(* IEC 61131-3 sources: BODAS-RC27-18_40/st/bodas_rc18_12_27_18_40/plc_logic/application/dsm_easyconfig/structure (part 2) *)

(* ---- dfc_rbr_ina57or-DFC_rbr_inA57OR.st ---- *)
(* --- Interface --- *)
{attribute 'external_name' := 'cmp_rts_DFC_rbr_inA57OR'}
TYPE DFC_rbr_inA57OR :
STRUCT
	DTC: UDINT := 16#134C00;
	DFCid: UINT := 81;
	debounceMethod: USINT := TIME_UP_DOWN;
END_STRUCT
END_TYPE

(* ---- dfc_rbr_ina57scb-DFC_rbr_inA57SCB.st ---- *)
(* --- Interface --- *)
{attribute 'external_name' := 'cmp_rts_DFC_rbr_inA57SCB'}
TYPE DFC_rbr_inA57SCB :
STRUCT
	DTC: UDINT := 16#134D00;
	DFCid: UINT := 82;
	debounceMethod: USINT := TIME_UP_DOWN;
END_STRUCT
END_TYPE

(* ---- dfc_rbr_ina57scg-DFC_rbr_inA57SCG.st ---- *)
(* --- Interface --- *)
{attribute 'external_name' := 'cmp_rts_DFC_rbr_inA57SCG'}
TYPE DFC_rbr_inA57SCG :
STRUCT
	DTC: UDINT := 16#134E00;
	DFCid: UINT := 83;
	debounceMethod: USINT := TIME_UP_DOWN;
END_STRUCT
END_TYPE

(* ---- dfc_rbr_ina59ol-DFC_rbr_inA59OL.st ---- *)
(* --- Interface --- *)
{attribute 'external_name' := 'cmp_rts_DFC_rbr_inA59OL'}
TYPE DFC_rbr_inA59OL :
STRUCT
	DTC: UDINT := 16#134F00;
	DFCid: UINT := 84;
	debounceMethod: USINT := TIME_UP_DOWN;
END_STRUCT
END_TYPE

(* ---- dfc_rbr_ina59scb-DFC_rbr_inA59SCB.st ---- *)
(* --- Interface --- *)
{attribute 'external_name' := 'cmp_rts_DFC_rbr_inA59SCB'}
TYPE DFC_rbr_inA59SCB :
STRUCT
	DTC: UDINT := 16#135000;
	DFCid: UINT := 85;
	debounceMethod: USINT := TIME_UP_DOWN;
END_STRUCT
END_TYPE

(* ---- dfc_rbr_ina59scg-DFC_rbr_inA59SCG.st ---- *)
(* --- Interface --- *)
{attribute 'external_name' := 'cmp_rts_DFC_rbr_inA59SCG'}
TYPE DFC_rbr_inA59SCG :
STRUCT
	DTC: UDINT := 16#135100;
	DFCid: UINT := 86;
	debounceMethod: USINT := TIME_UP_DOWN;
END_STRUCT
END_TYPE

(* ---- dfc_rbr_inai-DFC_rbr_inAi.st ---- *)
(* --- Interface --- *)
{attribute 'external_name' := 'cmp_rts_DFC_rbr_inAi'}
TYPE DFC_rbr_inAi :
STRUCT
	DTC: UDINT := 16#038000;
	DFCid: UINT := 578;
	debounceMethod: USINT := NO_DEBOUNCE;
END_STRUCT
END_TYPE

(* ---- dfc_rbr_inaic-DFC_rbr_inAic.st ---- *)
(* --- Interface --- *)
{attribute 'external_name' := 'cmp_rts_DFC_rbr_inAic'}
TYPE DFC_rbr_inAic :
STRUCT
	DTC: UDINT := 16#038100;
	DFCid: UINT := 579;
	debounceMethod: USINT := NO_DEBOUNCE;
END_STRUCT
END_TYPE

(* ---- dfc_rbr_inaiccfg-DFC_rbr_inAicCfg.st ---- *)
(* --- Interface --- *)
{attribute 'external_name' := 'cmp_rts_DFC_rbr_inAicCfg'}
TYPE DFC_rbr_inAicCfg :
STRUCT
	DTC: UDINT := 16#038200;
	DFCid: UINT := 580;
	debounceMethod: USINT := NO_DEBOUNCE;
END_STRUCT
END_TYPE

(* ---- dfc_rbr_inaicgetstatus-DFC_rbr_inAicGetStatus.st ---- *)
(* --- Interface --- *)
{attribute 'external_name' := 'cmp_rts_DFC_rbr_inAicGetStatus'}
TYPE DFC_rbr_inAicGetStatus :
STRUCT
	DTC: UDINT := 16#038D00;
	DFCid: UINT := 581;
	debounceMethod: USINT := NO_DEBOUNCE;
END_STRUCT
END_TYPE

(* ---- dfc_rbr_inaid-DFC_rbr_inAid.st ---- *)
(* --- Interface --- *)
{attribute 'external_name' := 'cmp_rts_DFC_rbr_inAid'}
TYPE DFC_rbr_inAid :
STRUCT
	DTC: UDINT := 16#038300;
	DFCid: UINT := 582;
	debounceMethod: USINT := NO_DEBOUNCE;
END_STRUCT
END_TYPE

(* ---- dfc_rbr_inaidcfg-DFC_rbr_inAidCfg.st ---- *)
(* --- Interface --- *)
{attribute 'external_name' := 'cmp_rts_DFC_rbr_inAidCfg'}
TYPE DFC_rbr_inAidCfg :
STRUCT
	DTC: UDINT := 16#038400;
	DFCid: UINT := 583;
	debounceMethod: USINT := NO_DEBOUNCE;
END_STRUCT
END_TYPE

(* ---- dfc_rbr_inaiv-DFC_rbr_inAiv.st ---- *)
(* --- Interface --- *)
{attribute 'external_name' := 'cmp_rts_DFC_rbr_inAiv'}
TYPE DFC_rbr_inAiv :
STRUCT
	DTC: UDINT := 16#038500;
	DFCid: UINT := 584;
	debounceMethod: USINT := NO_DEBOUNCE;
END_STRUCT
END_TYPE

(* ---- dfc_rbr_inaivcfg-DFC_rbr_inAivCfg.st ---- *)
(* --- Interface --- *)
{attribute 'external_name' := 'cmp_rts_DFC_rbr_inAivCfg'}
TYPE DFC_rbr_inAivCfg :
STRUCT
	DTC: UDINT := 16#038600;
	DFCid: UINT := 585;
	debounceMethod: USINT := NO_DEBOUNCE;
END_STRUCT
END_TYPE

(* ---- dfc_rbr_inaivgetstatus-DFC_rbr_inAivGetStatus.st ---- *)
(* --- Interface --- *)
{attribute 'external_name' := 'cmp_rts_DFC_rbr_inAivGetStatus'}
TYPE DFC_rbr_inAivGetStatus :
STRUCT
	DTC: UDINT := 16#038C00;
	DFCid: UINT := 586;
	debounceMethod: USINT := NO_DEBOUNCE;
END_STRUCT
END_TYPE

(* ---- dfc_rbr_indi-DFC_rbr_inDi.st ---- *)
(* --- Interface --- *)
{attribute 'external_name' := 'cmp_rts_DFC_rbr_inDi'}
TYPE DFC_rbr_inDi :
STRUCT
	DTC: UDINT := 16#038700;
	DFCid: UINT := 587;
	debounceMethod: USINT := NO_DEBOUNCE;
END_STRUCT
END_TYPE

(* ---- dfc_rbr_infi-DFC_rbr_inFi.st ---- *)
(* --- Interface --- *)
{attribute 'external_name' := 'cmp_rts_DFC_rbr_inFi'}
TYPE DFC_rbr_inFi :
STRUCT
	DTC: UDINT := 16#038800;
	DFCid: UINT := 588;
	debounceMethod: USINT := NO_DEBOUNCE;
END_STRUCT
END_TYPE

(* ---- dfc_rbr_infi_buffered-DFC_rbr_inFi_Buffered.st ---- *)
(* --- Interface --- *)
{attribute 'external_name' := 'cmp_rts_DFC_rbr_inFi_Buffered'}
TYPE DFC_rbr_inFi_Buffered :
STRUCT
	DTC: UDINT := 16#135200;
	DFCid: UINT := 591;
	debounceMethod: USINT := NO_DEBOUNCE;
END_STRUCT
END_TYPE

(* ---- dfc_rbr_inficfg-DFC_rbr_inFiCfg.st ---- *)
(* --- Interface --- *)
{attribute 'external_name' := 'cmp_rts_DFC_rbr_inFiCfg'}
TYPE DFC_rbr_inFiCfg :
STRUCT
	DTC: UDINT := 16#038900;
	DFCid: UINT := 589;
	debounceMethod: USINT := NO_DEBOUNCE;
END_STRUCT
END_TYPE

(* ---- dfc_rbr_infigetstatus-DFC_rbr_inFiGetStatus.st ---- *)
(* --- Interface --- *)
{attribute 'external_name' := 'cmp_rts_DFC_rbr_inFiGetStatus'}
TYPE DFC_rbr_inFiGetStatus :
STRUCT
	DTC: UDINT := 16#038F00;
	DFCid: UINT := 590;
	debounceMethod: USINT := NO_DEBOUNCE;
END_STRUCT
END_TYPE

(* ---- dfc_rbr_ink10or-DFC_rbr_inK10OR.st ---- *)
(* --- Interface --- *)
{attribute 'external_name' := 'cmp_rts_DFC_rbr_inK10OR'}
TYPE DFC_rbr_inK10OR :
STRUCT
	DTC: UDINT := 16#030100;
	DFCid: UINT := 87;
	debounceMethod: USINT := TIME_UP_DOWN;
END_STRUCT
END_TYPE

(* ---- dfc_rbr_ink10scb-DFC_rbr_inK10SCB.st ---- *)
(* --- Interface --- *)
{attribute 'external_name' := 'cmp_rts_DFC_rbr_inK10SCB'}
TYPE DFC_rbr_inK10SCB :
STRUCT
	DTC: UDINT := 16#030200;
	DFCid: UINT := 88;
	debounceMethod: USINT := TIME_UP_DOWN;
END_STRUCT
END_TYPE

(* ---- dfc_rbr_ink10scg-DFC_rbr_inK10SCG.st ---- *)
(* --- Interface --- *)
{attribute 'external_name' := 'cmp_rts_DFC_rbr_inK10SCG'}
TYPE DFC_rbr_inK10SCG :
STRUCT
	DTC: UDINT := 16#030300;
	DFCid: UINT := 89;
	debounceMethod: USINT := TIME_UP_DOWN;
END_STRUCT
END_TYPE

(* ---- dfc_rbr_ink11or-DFC_rbr_inK11OR.st ---- *)
(* --- Interface --- *)
{attribute 'external_name' := 'cmp_rts_DFC_rbr_inK11OR'}
TYPE DFC_rbr_inK11OR :
STRUCT
	DTC: UDINT := 16#03A200;
	DFCid: UINT := 90;
	debounceMethod: USINT := TIME_UP_DOWN;
END_STRUCT
END_TYPE

(* ---- dfc_rbr_ink11scb-DFC_rbr_inK11SCB.st ---- *)
(* --- Interface --- *)
{attribute 'external_name' := 'cmp_rts_DFC_rbr_inK11SCB'}
TYPE DFC_rbr_inK11SCB :
STRUCT
	DTC: UDINT := 16#03A300;
	DFCid: UINT := 91;
	debounceMethod: USINT := TIME_UP_DOWN;
END_STRUCT
END_TYPE

(* ---- dfc_rbr_ink11scg-DFC_rbr_inK11SCG.st ---- *)
(* --- Interface --- *)
{attribute 'external_name' := 'cmp_rts_DFC_rbr_inK11SCG'}
TYPE DFC_rbr_inK11SCG :
STRUCT
	DTC: UDINT := 16#03A400;
	DFCid: UINT := 92;
	debounceMethod: USINT := TIME_UP_DOWN;
END_STRUCT
END_TYPE

(* ---- dfc_rbr_ink30aicscb-DFC_rbr_inK30AicSCB.st ---- *)
(* --- Interface --- *)
{attribute 'external_name' := 'cmp_rts_DFC_rbr_inK30AicSCB'}
TYPE DFC_rbr_inK30AicSCB :
STRUCT
	DTC: UDINT := 16#03A500;
	DFCid: UINT := 93;
	debounceMethod: USINT := TIME_UP_DOWN;
END_STRUCT
END_TYPE

(* ---- dfc_rbr_ink30aicscg-DFC_rbr_inK30AicSCG.st ---- *)
(* --- Interface --- *)
{attribute 'external_name' := 'cmp_rts_DFC_rbr_inK30AicSCG'}
TYPE DFC_rbr_inK30AicSCG :
STRUCT
	DTC: UDINT := 16#03A600;
	DFCid: UINT := 94;
	debounceMethod: USINT := TIME_UP_DOWN;
END_STRUCT
END_TYPE

(* ---- dfc_rbr_ink30or-DFC_rbr_inK30OR.st ---- *)
(* --- Interface --- *)
{attribute 'external_name' := 'cmp_rts_DFC_rbr_inK30OR'}
TYPE DFC_rbr_inK30OR :
STRUCT
	DTC: UDINT := 16#03A700;
	DFCid: UINT := 95;
	debounceMethod: USINT := TIME_UP_DOWN;
END_STRUCT
END_TYPE

(* ---- dfc_rbr_ink30scb-DFC_rbr_inK30SCB.st ---- *)
(* --- Interface --- *)
{attribute 'external_name' := 'cmp_rts_DFC_rbr_inK30SCB'}
TYPE DFC_rbr_inK30SCB :
STRUCT
	DTC: UDINT := 16#03A800;
	DFCid: UINT := 96;
	debounceMethod: USINT := TIME_UP_DOWN;
END_STRUCT
END_TYPE

(* ---- dfc_rbr_ink30scg-DFC_rbr_inK30SCG.st ---- *)
(* --- Interface --- *)
{attribute 'external_name' := 'cmp_rts_DFC_rbr_inK30SCG'}
TYPE DFC_rbr_inK30SCG :
STRUCT
	DTC: UDINT := 16#03A900;
	DFCid: UINT := 97;
	debounceMethod: USINT := TIME_UP_DOWN;
END_STRUCT
END_TYPE

(* ---- dfc_rbr_ink30shuntscb-DFC_rbr_inK30ShuntSCB.st ---- *)
(* --- Interface --- *)
{attribute 'external_name' := 'cmp_rts_DFC_rbr_inK30ShuntSCB'}
TYPE DFC_rbr_inK30ShuntSCB :
STRUCT
	DTC: UDINT := 16#03AA00;
	DFCid: UINT := 98;
	debounceMethod: USINT := TIME_UP_DOWN;
END_STRUCT
END_TYPE

(* ---- dfc_rbr_ink31or-DFC_rbr_inK31OR.st ---- *)
(* --- Interface --- *)
{attribute 'external_name' := 'cmp_rts_DFC_rbr_inK31OR'}
TYPE DFC_rbr_inK31OR :
STRUCT
	DTC: UDINT := 16#03AB00;
	DFCid: UINT := 99;
	debounceMethod: USINT := TIME_UP_DOWN;
END_STRUCT
END_TYPE

(* ---- dfc_rbr_ink31scb-DFC_rbr_inK31SCB.st ---- *)
(* --- Interface --- *)
{attribute 'external_name' := 'cmp_rts_DFC_rbr_inK31SCB'}
TYPE DFC_rbr_inK31SCB :
STRUCT
	DTC: UDINT := 16#03AC00;
	DFCid: UINT := 100;
	debounceMethod: USINT := TIME_UP_DOWN;
END_STRUCT
END_TYPE

(* ---- dfc_rbr_ink31scg-DFC_rbr_inK31SCG.st ---- *)
(* --- Interface --- *)
{attribute 'external_name' := 'cmp_rts_DFC_rbr_inK31SCG'}
TYPE DFC_rbr_inK31SCG :
STRUCT
	DTC: UDINT := 16#03AD00;
	DFCid: UINT := 101;
	debounceMethod: USINT := TIME_UP_DOWN;
END_STRUCT
END_TYPE

(* ---- dfc_rbr_ink32or-DFC_rbr_inK32OR.st ---- *)
(* --- Interface --- *)
{attribute 'external_name' := 'cmp_rts_DFC_rbr_inK32OR'}
TYPE DFC_rbr_inK32OR :
STRUCT
	DTC: UDINT := 16#03AE00;
	DFCid: UINT := 102;
	debounceMethod: USINT := TIME_UP_DOWN;
END_STRUCT
END_TYPE

(* ---- dfc_rbr_ink32scb-DFC_rbr_inK32SCB.st ---- *)
(* --- Interface --- *)
{attribute 'external_name' := 'cmp_rts_DFC_rbr_inK32SCB'}
TYPE DFC_rbr_inK32SCB :
STRUCT
	DTC: UDINT := 16#03AF00;
	DFCid: UINT := 103;
	debounceMethod: USINT := TIME_UP_DOWN;
END_STRUCT
END_TYPE

(* ---- dfc_rbr_ink32scg-DFC_rbr_inK32SCG.st ---- *)
(* --- Interface --- *)
{attribute 'external_name' := 'cmp_rts_DFC_rbr_inK32SCG'}
TYPE DFC_rbr_inK32SCG :
STRUCT
	DTC: UDINT := 16#03B000;
	DFCid: UINT := 104;
	debounceMethod: USINT := TIME_UP_DOWN;
END_STRUCT
END_TYPE

(* ---- dfc_rbr_ink33or-DFC_rbr_inK33OR.st ---- *)
(* --- Interface --- *)
{attribute 'external_name' := 'cmp_rts_DFC_rbr_inK33OR'}
TYPE DFC_rbr_inK33OR :
STRUCT
	DTC: UDINT := 16#03B100;
	DFCid: UINT := 105;
	debounceMethod: USINT := TIME_UP_DOWN;
END_STRUCT
END_TYPE

(* ---- dfc_rbr_ink33scb-DFC_rbr_inK33SCB.st ---- *)
(* --- Interface --- *)
{attribute 'external_name' := 'cmp_rts_DFC_rbr_inK33SCB'}
TYPE DFC_rbr_inK33SCB :
STRUCT
	DTC: UDINT := 16#03B200;
	DFCid: UINT := 106;
	debounceMethod: USINT := TIME_UP_DOWN;
END_STRUCT
END_TYPE

(* ---- dfc_rbr_ink33scg-DFC_rbr_inK33SCG.st ---- *)
(* --- Interface --- *)
{attribute 'external_name' := 'cmp_rts_DFC_rbr_inK33SCG'}
TYPE DFC_rbr_inK33SCG :
STRUCT
	DTC: UDINT := 16#03B300;
	DFCid: UINT := 107;
	debounceMethod: USINT := TIME_UP_DOWN;
END_STRUCT
END_TYPE

(* ---- dfc_rbr_ink34or-DFC_rbr_inK34OR.st ---- *)
(* --- Interface --- *)
{attribute 'external_name' := 'cmp_rts_DFC_rbr_inK34OR'}
TYPE DFC_rbr_inK34OR :
STRUCT
	DTC: UDINT := 16#03B400;
	DFCid: UINT := 108;
	debounceMethod: USINT := TIME_UP_DOWN;
END_STRUCT
END_TYPE

(* ---- dfc_rbr_ink34scb-DFC_rbr_inK34SCB.st ---- *)
(* --- Interface --- *)
{attribute 'external_name' := 'cmp_rts_DFC_rbr_inK34SCB'}
TYPE DFC_rbr_inK34SCB :
STRUCT
	DTC: UDINT := 16#03B500;
	DFCid: UINT := 109;
	debounceMethod: USINT := TIME_UP_DOWN;
END_STRUCT
END_TYPE

(* ---- dfc_rbr_ink34scg-DFC_rbr_inK34SCG.st ---- *)
(* --- Interface --- *)
{attribute 'external_name' := 'cmp_rts_DFC_rbr_inK34SCG'}
TYPE DFC_rbr_inK34SCG :
STRUCT
	DTC: UDINT := 16#03B600;
	DFCid: UINT := 110;
	debounceMethod: USINT := TIME_UP_DOWN;
END_STRUCT
END_TYPE

(* ---- dfc_rbr_ink35or-DFC_rbr_inK35OR.st ---- *)
(* --- Interface --- *)
{attribute 'external_name' := 'cmp_rts_DFC_rbr_inK35OR'}
TYPE DFC_rbr_inK35OR :
STRUCT
	DTC: UDINT := 16#03B700;
	DFCid: UINT := 111;
	debounceMethod: USINT := TIME_UP_DOWN;
END_STRUCT
END_TYPE

(* ---- dfc_rbr_ink35scb-DFC_rbr_inK35SCB.st ---- *)
(* --- Interface --- *)
{attribute 'external_name' := 'cmp_rts_DFC_rbr_inK35SCB'}
TYPE DFC_rbr_inK35SCB :
STRUCT
	DTC: UDINT := 16#03B800;
	DFCid: UINT := 112;
	debounceMethod: USINT := TIME_UP_DOWN;
END_STRUCT
END_TYPE

(* ---- dfc_rbr_ink35scg-DFC_rbr_inK35SCG.st ---- *)
(* --- Interface --- *)
{attribute 'external_name' := 'cmp_rts_DFC_rbr_inK35SCG'}
TYPE DFC_rbr_inK35SCG :
STRUCT
	DTC: UDINT := 16#03B900;
	DFCid: UINT := 113;
	debounceMethod: USINT := TIME_UP_DOWN;
END_STRUCT
END_TYPE

(* ---- dfc_rbr_ink36or-DFC_rbr_inK36OR.st ---- *)
(* --- Interface --- *)
{attribute 'external_name' := 'cmp_rts_DFC_rbr_inK36OR'}
TYPE DFC_rbr_inK36OR :
STRUCT
	DTC: UDINT := 16#030400;
	DFCid: UINT := 114;
	debounceMethod: USINT := TIME_UP_DOWN;
END_STRUCT
END_TYPE

(* ---- dfc_rbr_ink36scb-DFC_rbr_inK36SCB.st ---- *)
(* --- Interface --- *)
{attribute 'external_name' := 'cmp_rts_DFC_rbr_inK36SCB'}
TYPE DFC_rbr_inK36SCB :
STRUCT
	DTC: UDINT := 16#030500;
	DFCid: UINT := 115;
	debounceMethod: USINT := TIME_UP_DOWN;
END_STRUCT
END_TYPE

(* ---- dfc_rbr_ink36scg-DFC_rbr_inK36SCG.st ---- *)
(* --- Interface --- *)
{attribute 'external_name' := 'cmp_rts_DFC_rbr_inK36SCG'}
TYPE DFC_rbr_inK36SCG :
STRUCT
	DTC: UDINT := 16#030600;
	DFCid: UINT := 116;
	debounceMethod: USINT := TIME_UP_DOWN;
END_STRUCT
END_TYPE

(* ---- dfc_rbr_ink37aicscb-DFC_rbr_inK37AicSCB.st ---- *)
(* --- Interface --- *)
{attribute 'external_name' := 'cmp_rts_DFC_rbr_inK37AicSCB'}
TYPE DFC_rbr_inK37AicSCB :
STRUCT
	DTC: UDINT := 16#030700;
	DFCid: UINT := 117;
	debounceMethod: USINT := TIME_UP_DOWN;
END_STRUCT
END_TYPE

(* ---- dfc_rbr_ink37aicscg-DFC_rbr_inK37AicSCG.st ---- *)
(* --- Interface --- *)
{attribute 'external_name' := 'cmp_rts_DFC_rbr_inK37AicSCG'}
TYPE DFC_rbr_inK37AicSCG :
STRUCT
	DTC: UDINT := 16#030800;
	DFCid: UINT := 118;
	debounceMethod: USINT := TIME_UP_DOWN;
END_STRUCT
END_TYPE

(* ---- dfc_rbr_ink37or-DFC_rbr_inK37OR.st ---- *)
(* --- Interface --- *)
{attribute 'external_name' := 'cmp_rts_DFC_rbr_inK37OR'}
TYPE DFC_rbr_inK37OR :
STRUCT
	DTC: UDINT := 16#030900;
	DFCid: UINT := 119;
	debounceMethod: USINT := TIME_UP_DOWN;
END_STRUCT
END_TYPE

(* ---- dfc_rbr_ink37scb-DFC_rbr_inK37SCB.st ---- *)
(* --- Interface --- *)
{attribute 'external_name' := 'cmp_rts_DFC_rbr_inK37SCB'}
TYPE DFC_rbr_inK37SCB :
STRUCT
	DTC: UDINT := 16#030A00;
	DFCid: UINT := 120;
	debounceMethod: USINT := TIME_UP_DOWN;
END_STRUCT
END_TYPE

(* ---- dfc_rbr_ink37scg-DFC_rbr_inK37SCG.st ---- *)
(* --- Interface --- *)
{attribute 'external_name' := 'cmp_rts_DFC_rbr_inK37SCG'}
TYPE DFC_rbr_inK37SCG :
STRUCT
	DTC: UDINT := 16#030B00;
	DFCid: UINT := 121;
	debounceMethod: USINT := TIME_UP_DOWN;
END_STRUCT
END_TYPE

(* ---- dfc_rbr_ink37shuntscb-DFC_rbr_inK37ShuntSCB.st ---- *)
(* --- Interface --- *)
{attribute 'external_name' := 'cmp_rts_DFC_rbr_inK37ShuntSCB'}
TYPE DFC_rbr_inK37ShuntSCB :
STRUCT
	DTC: UDINT := 16#030C00;
	DFCid: UINT := 122;
	debounceMethod: USINT := TIME_UP_DOWN;
END_STRUCT
END_TYPE

(* ---- dfc_rbr_ink38aicscb-DFC_rbr_inK38AicSCB.st ---- *)
(* --- Interface --- *)
{attribute 'external_name' := 'cmp_rts_DFC_rbr_inK38AicSCB'}
TYPE DFC_rbr_inK38AicSCB :
STRUCT
	DTC: UDINT := 16#03BA00;
	DFCid: UINT := 123;
	debounceMethod: USINT := TIME_UP_DOWN;
END_STRUCT
END_TYPE

(* ---- dfc_rbr_ink38aicscg-DFC_rbr_inK38AicSCG.st ---- *)
(* --- Interface --- *)
{attribute 'external_name' := 'cmp_rts_DFC_rbr_inK38AicSCG'}
TYPE DFC_rbr_inK38AicSCG :
STRUCT
	DTC: UDINT := 16#03BB00;
	DFCid: UINT := 124;
	debounceMethod: USINT := TIME_UP_DOWN;
END_STRUCT
END_TYPE

(* ---- dfc_rbr_ink38or-DFC_rbr_inK38OR.st ---- *)
(* --- Interface --- *)
{attribute 'external_name' := 'cmp_rts_DFC_rbr_inK38OR'}
TYPE DFC_rbr_inK38OR :
STRUCT
	DTC: UDINT := 16#030D00;
	DFCid: UINT := 125;
	debounceMethod: USINT := TIME_UP_DOWN;
END_STRUCT
END_TYPE

(* ---- dfc_rbr_ink38scb-DFC_rbr_inK38SCB.st ---- *)
(* --- Interface --- *)
{attribute 'external_name' := 'cmp_rts_DFC_rbr_inK38SCB'}
TYPE DFC_rbr_inK38SCB :
STRUCT
	DTC: UDINT := 16#030E00;
	DFCid: UINT := 126;
	debounceMethod: USINT := TIME_UP_DOWN;
END_STRUCT
END_TYPE

(* ---- dfc_rbr_ink38scg-DFC_rbr_inK38SCG.st ---- *)
(* --- Interface --- *)
{attribute 'external_name' := 'cmp_rts_DFC_rbr_inK38SCG'}
TYPE DFC_rbr_inK38SCG :
STRUCT
	DTC: UDINT := 16#030F00;
	DFCid: UINT := 127;
	debounceMethod: USINT := TIME_UP_DOWN;
END_STRUCT
END_TYPE

(* ---- dfc_rbr_ink38shuntscb-DFC_rbr_inK38ShuntSCB.st ---- *)
(* --- Interface --- *)
{attribute 'external_name' := 'cmp_rts_DFC_rbr_inK38ShuntSCB'}
TYPE DFC_rbr_inK38ShuntSCB :
STRUCT
	DTC: UDINT := 16#03BC00;
	DFCid: UINT := 128;
	debounceMethod: USINT := TIME_UP_DOWN;
END_STRUCT
END_TYPE

(* ---- dfc_rbr_ink39aicscb-DFC_rbr_inK39AicSCB.st ---- *)
(* --- Interface --- *)
{attribute 'external_name' := 'cmp_rts_DFC_rbr_inK39AicSCB'}
TYPE DFC_rbr_inK39AicSCB :
STRUCT
	DTC: UDINT := 16#03BD00;
	DFCid: UINT := 129;
	debounceMethod: USINT := TIME_UP_DOWN;
END_STRUCT
END_TYPE

(* ---- dfc_rbr_ink39aicscg-DFC_rbr_inK39AicSCG.st ---- *)
(* --- Interface --- *)
{attribute 'external_name' := 'cmp_rts_DFC_rbr_inK39AicSCG'}
TYPE DFC_rbr_inK39AicSCG :
STRUCT
	DTC: UDINT := 16#03BE00;
	DFCid: UINT := 130;
	debounceMethod: USINT := TIME_UP_DOWN;
END_STRUCT
END_TYPE

(* ---- dfc_rbr_ink39or-DFC_rbr_inK39OR.st ---- *)
(* --- Interface --- *)
{attribute 'external_name' := 'cmp_rts_DFC_rbr_inK39OR'}
TYPE DFC_rbr_inK39OR :
STRUCT
	DTC: UDINT := 16#031000;
	DFCid: UINT := 131;
	debounceMethod: USINT := TIME_UP_DOWN;
END_STRUCT
END_TYPE

(* ---- dfc_rbr_ink39scb-DFC_rbr_inK39SCB.st ---- *)
(* --- Interface --- *)
{attribute 'external_name' := 'cmp_rts_DFC_rbr_inK39SCB'}
TYPE DFC_rbr_inK39SCB :
STRUCT
	DTC: UDINT := 16#031100;
	DFCid: UINT := 132;
	debounceMethod: USINT := TIME_UP_DOWN;
END_STRUCT
END_TYPE

(* ---- dfc_rbr_ink39scg-DFC_rbr_inK39SCG.st ---- *)
(* --- Interface --- *)
{attribute 'external_name' := 'cmp_rts_DFC_rbr_inK39SCG'}
TYPE DFC_rbr_inK39SCG :
STRUCT
	DTC: UDINT := 16#031200;
	DFCid: UINT := 133;
	debounceMethod: USINT := TIME_UP_DOWN;
END_STRUCT
END_TYPE

(* ---- dfc_rbr_ink39shuntscb-DFC_rbr_inK39ShuntSCB.st ---- *)
(* --- Interface --- *)
{attribute 'external_name' := 'cmp_rts_DFC_rbr_inK39ShuntSCB'}
TYPE DFC_rbr_inK39ShuntSCB :
STRUCT
	DTC: UDINT := 16#03BF00;
	DFCid: UINT := 134;
	debounceMethod: USINT := TIME_UP_DOWN;
END_STRUCT
END_TYPE

(* ---- dfc_rbr_ink40aicscb-DFC_rbr_inK40AicSCB.st ---- *)
(* --- Interface --- *)
{attribute 'external_name' := 'cmp_rts_DFC_rbr_inK40AicSCB'}
TYPE DFC_rbr_inK40AicSCB :
STRUCT
	DTC: UDINT := 16#03C000;
	DFCid: UINT := 135;
	debounceMethod: USINT := TIME_UP_DOWN;
END_STRUCT
END_TYPE

(* ---- dfc_rbr_ink40aicscg-DFC_rbr_inK40AicSCG.st ---- *)
(* --- Interface --- *)
{attribute 'external_name' := 'cmp_rts_DFC_rbr_inK40AicSCG'}
TYPE DFC_rbr_inK40AicSCG :
STRUCT
	DTC: UDINT := 16#03C100;
	DFCid: UINT := 136;
	debounceMethod: USINT := TIME_UP_DOWN;
END_STRUCT
END_TYPE

(* ---- dfc_rbr_ink40or-DFC_rbr_inK40OR.st ---- *)
(* --- Interface --- *)
{attribute 'external_name' := 'cmp_rts_DFC_rbr_inK40OR'}
TYPE DFC_rbr_inK40OR :
STRUCT
	DTC: UDINT := 16#031300;
	DFCid: UINT := 137;
	debounceMethod: USINT := TIME_UP_DOWN;
END_STRUCT
END_TYPE

(* ---- dfc_rbr_ink40scb-DFC_rbr_inK40SCB.st ---- *)
(* --- Interface --- *)
{attribute 'external_name' := 'cmp_rts_DFC_rbr_inK40SCB'}
TYPE DFC_rbr_inK40SCB :
STRUCT
	DTC: UDINT := 16#031400;
	DFCid: UINT := 138;
	debounceMethod: USINT := TIME_UP_DOWN;
END_STRUCT
END_TYPE

(* ---- dfc_rbr_ink40scg-DFC_rbr_inK40SCG.st ---- *)
(* --- Interface --- *)
{attribute 'external_name' := 'cmp_rts_DFC_rbr_inK40SCG'}
TYPE DFC_rbr_inK40SCG :
STRUCT
	DTC: UDINT := 16#031500;
	DFCid: UINT := 139;
	debounceMethod: USINT := TIME_UP_DOWN;
END_STRUCT
END_TYPE

(* ---- dfc_rbr_ink40shuntscb-DFC_rbr_inK40ShuntSCB.st ---- *)
(* --- Interface --- *)
{attribute 'external_name' := 'cmp_rts_DFC_rbr_inK40ShuntSCB'}
TYPE DFC_rbr_inK40ShuntSCB :
STRUCT
	DTC: UDINT := 16#03C200;
	DFCid: UINT := 140;
	debounceMethod: USINT := TIME_UP_DOWN;
END_STRUCT
END_TYPE

(* ---- dfc_rbr_ink41aicscb-DFC_rbr_inK41AicSCB.st ---- *)
(* --- Interface --- *)
{attribute 'external_name' := 'cmp_rts_DFC_rbr_inK41AicSCB'}
TYPE DFC_rbr_inK41AicSCB :
STRUCT
	DTC: UDINT := 16#03C300;
	DFCid: UINT := 141;
	debounceMethod: USINT := TIME_UP_DOWN;
END_STRUCT
END_TYPE

(* ---- dfc_rbr_ink41aicscg-DFC_rbr_inK41AicSCG.st ---- *)
(* --- Interface --- *)
{attribute 'external_name' := 'cmp_rts_DFC_rbr_inK41AicSCG'}
TYPE DFC_rbr_inK41AicSCG :
STRUCT
	DTC: UDINT := 16#03C400;
	DFCid: UINT := 142;
	debounceMethod: USINT := TIME_UP_DOWN;
END_STRUCT
END_TYPE

(* ---- dfc_rbr_ink41or-DFC_rbr_inK41OR.st ---- *)
(* --- Interface --- *)
{attribute 'external_name' := 'cmp_rts_DFC_rbr_inK41OR'}
TYPE DFC_rbr_inK41OR :
STRUCT
	DTC: UDINT := 16#031600;
	DFCid: UINT := 143;
	debounceMethod: USINT := TIME_UP_DOWN;
END_STRUCT
END_TYPE

(* ---- dfc_rbr_ink41scb-DFC_rbr_inK41SCB.st ---- *)
(* --- Interface --- *)
{attribute 'external_name' := 'cmp_rts_DFC_rbr_inK41SCB'}
TYPE DFC_rbr_inK41SCB :
STRUCT
	DTC: UDINT := 16#031700;
	DFCid: UINT := 144;
	debounceMethod: USINT := TIME_UP_DOWN;
END_STRUCT
END_TYPE

(* ---- dfc_rbr_ink41scg-DFC_rbr_inK41SCG.st ---- *)
(* --- Interface --- *)
{attribute 'external_name' := 'cmp_rts_DFC_rbr_inK41SCG'}
TYPE DFC_rbr_inK41SCG :
STRUCT
	DTC: UDINT := 16#031800;
	DFCid: UINT := 145;
	debounceMethod: USINT := TIME_UP_DOWN;
END_STRUCT
END_TYPE

(* ---- dfc_rbr_ink41shuntscb-DFC_rbr_inK41ShuntSCB.st ---- *)
(* --- Interface --- *)
{attribute 'external_name' := 'cmp_rts_DFC_rbr_inK41ShuntSCB'}
TYPE DFC_rbr_inK41ShuntSCB :
STRUCT
	DTC: UDINT := 16#03C500;
	DFCid: UINT := 146;
	debounceMethod: USINT := TIME_UP_DOWN;
END_STRUCT
END_TYPE

(* ---- dfc_rbr_ink42aicscb-DFC_rbr_inK42AicSCB.st ---- *)
(* --- Interface --- *)
{attribute 'external_name' := 'cmp_rts_DFC_rbr_inK42AicSCB'}
TYPE DFC_rbr_inK42AicSCB :
STRUCT
	DTC: UDINT := 16#03C600;
	DFCid: UINT := 147;
	debounceMethod: USINT := TIME_UP_DOWN;
END_STRUCT
END_TYPE

(* ---- dfc_rbr_ink42aicscg-DFC_rbr_inK42AicSCG.st ---- *)
(* --- Interface --- *)
{attribute 'external_name' := 'cmp_rts_DFC_rbr_inK42AicSCG'}
TYPE DFC_rbr_inK42AicSCG :
STRUCT
	DTC: UDINT := 16#03C700;
	DFCid: UINT := 148;
	debounceMethod: USINT := TIME_UP_DOWN;
END_STRUCT
END_TYPE

(* ---- dfc_rbr_ink42or-DFC_rbr_inK42OR.st ---- *)
(* --- Interface --- *)
{attribute 'external_name' := 'cmp_rts_DFC_rbr_inK42OR'}
TYPE DFC_rbr_inK42OR :
STRUCT
	DTC: UDINT := 16#031900;
	DFCid: UINT := 149;
	debounceMethod: USINT := TIME_UP_DOWN;
END_STRUCT
END_TYPE

(* ---- dfc_rbr_ink42scb-DFC_rbr_inK42SCB.st ---- *)
(* --- Interface --- *)
{attribute 'external_name' := 'cmp_rts_DFC_rbr_inK42SCB'}
TYPE DFC_rbr_inK42SCB :
STRUCT
	DTC: UDINT := 16#031A00;
	DFCid: UINT := 150;
	debounceMethod: USINT := TIME_UP_DOWN;
END_STRUCT
END_TYPE

(* ---- dfc_rbr_ink42scg-DFC_rbr_inK42SCG.st ---- *)
(* --- Interface --- *)
{attribute 'external_name' := 'cmp_rts_DFC_rbr_inK42SCG'}
TYPE DFC_rbr_inK42SCG :
STRUCT
	DTC: UDINT := 16#031B00;
	DFCid: UINT := 151;
	debounceMethod: USINT := TIME_UP_DOWN;
END_STRUCT
END_TYPE

(* ---- dfc_rbr_ink42shuntscb-DFC_rbr_inK42ShuntSCB.st ---- *)
(* --- Interface --- *)
{attribute 'external_name' := 'cmp_rts_DFC_rbr_inK42ShuntSCB'}
TYPE DFC_rbr_inK42ShuntSCB :
STRUCT
	DTC: UDINT := 16#03C800;
	DFCid: UINT := 152;
	debounceMethod: USINT := TIME_UP_DOWN;
END_STRUCT
END_TYPE

(* ---- dfc_rbr_ink43or-DFC_rbr_inK43OR.st ---- *)
(* --- Interface --- *)
{attribute 'external_name' := 'cmp_rts_DFC_rbr_inK43OR'}
TYPE DFC_rbr_inK43OR :
STRUCT
	DTC: UDINT := 16#031C00;
	DFCid: UINT := 153;
	debounceMethod: USINT := TIME_UP_DOWN;
END_STRUCT
END_TYPE

(* ---- dfc_rbr_ink43scb-DFC_rbr_inK43SCB.st ---- *)
(* --- Interface --- *)
{attribute 'external_name' := 'cmp_rts_DFC_rbr_inK43SCB'}
TYPE DFC_rbr_inK43SCB :
STRUCT
	DTC: UDINT := 16#031D00;
	DFCid: UINT := 154;
	debounceMethod: USINT := TIME_UP_DOWN;
END_STRUCT
END_TYPE

(* ---- dfc_rbr_ink43scg-DFC_rbr_inK43SCG.st ---- *)
(* --- Interface --- *)
{attribute 'external_name' := 'cmp_rts_DFC_rbr_inK43SCG'}
TYPE DFC_rbr_inK43SCG :
STRUCT
	DTC: UDINT := 16#031E00;
	DFCid: UINT := 155;
	debounceMethod: USINT := TIME_UP_DOWN;
END_STRUCT
END_TYPE

(* ---- dfc_rbr_ink44aicscb-DFC_rbr_inK44AicSCB.st ---- *)
(* --- Interface --- *)
{attribute 'external_name' := 'cmp_rts_DFC_rbr_inK44AicSCB'}
TYPE DFC_rbr_inK44AicSCB :
STRUCT
	DTC: UDINT := 16#03C900;
	DFCid: UINT := 156;
	debounceMethod: USINT := TIME_UP_DOWN;
END_STRUCT
END_TYPE

(* ---- dfc_rbr_ink44aicscg-DFC_rbr_inK44AicSCG.st ---- *)
(* --- Interface --- *)
{attribute 'external_name' := 'cmp_rts_DFC_rbr_inK44AicSCG'}
TYPE DFC_rbr_inK44AicSCG :
STRUCT
	DTC: UDINT := 16#03CA00;
	DFCid: UINT := 157;
	debounceMethod: USINT := TIME_UP_DOWN;
END_STRUCT
END_TYPE

(* ---- dfc_rbr_ink44or-DFC_rbr_inK44OR.st ---- *)
(* --- Interface --- *)
{attribute 'external_name' := 'cmp_rts_DFC_rbr_inK44OR'}
TYPE DFC_rbr_inK44OR :
STRUCT
	DTC: UDINT := 16#031F00;
	DFCid: UINT := 158;
	debounceMethod: USINT := TIME_UP_DOWN;
END_STRUCT
END_TYPE

(* ---- dfc_rbr_ink44scb-DFC_rbr_inK44SCB.st ---- *)
(* --- Interface --- *)
{attribute 'external_name' := 'cmp_rts_DFC_rbr_inK44SCB'}
TYPE DFC_rbr_inK44SCB :
STRUCT
	DTC: UDINT := 16#032000;
	DFCid: UINT := 159;
	debounceMethod: USINT := TIME_UP_DOWN;
END_STRUCT
END_TYPE

(* ---- dfc_rbr_ink44scg-DFC_rbr_inK44SCG.st ---- *)
(* --- Interface --- *)
{attribute 'external_name' := 'cmp_rts_DFC_rbr_inK44SCG'}
TYPE DFC_rbr_inK44SCG :
STRUCT
	DTC: UDINT := 16#032100;
	DFCid: UINT := 160;
	debounceMethod: USINT := TIME_UP_DOWN;
END_STRUCT
END_TYPE

(* ---- dfc_rbr_ink44shuntscb-DFC_rbr_inK44ShuntSCB.st ---- *)
(* --- Interface --- *)
{attribute 'external_name' := 'cmp_rts_DFC_rbr_inK44ShuntSCB'}
TYPE DFC_rbr_inK44ShuntSCB :
STRUCT
	DTC: UDINT := 16#03CB00;
	DFCid: UINT := 161;
	debounceMethod: USINT := TIME_UP_DOWN;
END_STRUCT
END_TYPE

(* ---- dfc_rbr_ink45aicscb-DFC_rbr_inK45AicSCB.st ---- *)
(* --- Interface --- *)
{attribute 'external_name' := 'cmp_rts_DFC_rbr_inK45AicSCB'}
TYPE DFC_rbr_inK45AicSCB :
STRUCT
	DTC: UDINT := 16#03CC00;
	DFCid: UINT := 162;
	debounceMethod: USINT := TIME_UP_DOWN;
END_STRUCT
END_TYPE

(* ---- dfc_rbr_ink45aicscg-DFC_rbr_inK45AicSCG.st ---- *)
(* --- Interface --- *)
{attribute 'external_name' := 'cmp_rts_DFC_rbr_inK45AicSCG'}
TYPE DFC_rbr_inK45AicSCG :
STRUCT
	DTC: UDINT := 16#03CD00;
	DFCid: UINT := 163;
	debounceMethod: USINT := TIME_UP_DOWN;
END_STRUCT
END_TYPE

(* ---- dfc_rbr_ink45or-DFC_rbr_inK45OR.st ---- *)
(* --- Interface --- *)
{attribute 'external_name' := 'cmp_rts_DFC_rbr_inK45OR'}
TYPE DFC_rbr_inK45OR :
STRUCT
	DTC: UDINT := 16#032200;
	DFCid: UINT := 164;
	debounceMethod: USINT := TIME_UP_DOWN;
END_STRUCT
END_TYPE

(* ---- dfc_rbr_ink45scb-DFC_rbr_inK45SCB.st ---- *)
(* --- Interface --- *)
{attribute 'external_name' := 'cmp_rts_DFC_rbr_inK45SCB'}
TYPE DFC_rbr_inK45SCB :
STRUCT
	DTC: UDINT := 16#032300;
	DFCid: UINT := 165;
	debounceMethod: USINT := TIME_UP_DOWN;
END_STRUCT
END_TYPE

(* ---- dfc_rbr_ink45scg-DFC_rbr_inK45SCG.st ---- *)
(* --- Interface --- *)
{attribute 'external_name' := 'cmp_rts_DFC_rbr_inK45SCG'}
TYPE DFC_rbr_inK45SCG :
STRUCT
	DTC: UDINT := 16#032400;
	DFCid: UINT := 166;
	debounceMethod: USINT := TIME_UP_DOWN;
END_STRUCT
END_TYPE

(* ---- dfc_rbr_ink45shuntscb-DFC_rbr_inK45ShuntSCB.st ---- *)
(* --- Interface --- *)
{attribute 'external_name' := 'cmp_rts_DFC_rbr_inK45ShuntSCB'}
TYPE DFC_rbr_inK45ShuntSCB :
STRUCT
	DTC: UDINT := 16#03CE00;
	DFCid: UINT := 167;
	debounceMethod: USINT := TIME_UP_DOWN;
END_STRUCT
END_TYPE

(* ---- dfc_rbr_ink52or-DFC_rbr_inK52OR.st ---- *)
(* --- Interface --- *)
{attribute 'external_name' := 'cmp_rts_DFC_rbr_inK52OR'}
TYPE DFC_rbr_inK52OR :
STRUCT
	DTC: UDINT := 16#032500;
	DFCid: UINT := 168;
	debounceMethod: USINT := TIME_UP_DOWN;
END_STRUCT
END_TYPE

(* ---- dfc_rbr_ink52scb-DFC_rbr_inK52SCB.st ---- *)
(* --- Interface --- *)
{attribute 'external_name' := 'cmp_rts_DFC_rbr_inK52SCB'}
TYPE DFC_rbr_inK52SCB :
STRUCT
	DTC: UDINT := 16#032600;
	DFCid: UINT := 169;
	debounceMethod: USINT := TIME_UP_DOWN;
END_STRUCT
END_TYPE

(* ---- dfc_rbr_ink52scg-DFC_rbr_inK52SCG.st ---- *)
(* --- Interface --- *)
{attribute 'external_name' := 'cmp_rts_DFC_rbr_inK52SCG'}
TYPE DFC_rbr_inK52SCG :
STRUCT
	DTC: UDINT := 16#032700;
	DFCid: UINT := 170;
	debounceMethod: USINT := TIME_UP_DOWN;
END_STRUCT
END_TYPE

(* ---- dfc_rbr_ink53or-DFC_rbr_inK53OR.st ---- *)
(* --- Interface --- *)
{attribute 'external_name' := 'cmp_rts_DFC_rbr_inK53OR'}
TYPE DFC_rbr_inK53OR :
STRUCT
	DTC: UDINT := 16#032800;
	DFCid: UINT := 171;
	debounceMethod: USINT := TIME_UP_DOWN;
END_STRUCT
END_TYPE

(* ---- dfc_rbr_ink53scb-DFC_rbr_inK53SCB.st ---- *)
(* --- Interface --- *)
{attribute 'external_name' := 'cmp_rts_DFC_rbr_inK53SCB'}
TYPE DFC_rbr_inK53SCB :
STRUCT
	DTC: UDINT := 16#032900;
	DFCid: UINT := 172;
	debounceMethod: USINT := TIME_UP_DOWN;
END_STRUCT
END_TYPE

(* ---- dfc_rbr_ink53scg-DFC_rbr_inK53SCG.st ---- *)
(* --- Interface --- *)
{attribute 'external_name' := 'cmp_rts_DFC_rbr_inK53SCG'}
TYPE DFC_rbr_inK53SCG :
STRUCT
	DTC: UDINT := 16#032A00;
	DFCid: UINT := 173;
	debounceMethod: USINT := TIME_UP_DOWN;
END_STRUCT
END_TYPE

(* ---- dfc_rbr_ink54aicscb-DFC_rbr_inK54AicSCB.st ---- *)
(* --- Interface --- *)
{attribute 'external_name' := 'cmp_rts_DFC_rbr_inK54AicSCB'}
TYPE DFC_rbr_inK54AicSCB :
STRUCT
	DTC: UDINT := 16#032B00;
	DFCid: UINT := 174;
	debounceMethod: USINT := TIME_UP_DOWN;
END_STRUCT
END_TYPE

(* ---- dfc_rbr_ink54aicscg-DFC_rbr_inK54AicSCG.st ---- *)
(* --- Interface --- *)
{attribute 'external_name' := 'cmp_rts_DFC_rbr_inK54AicSCG'}
TYPE DFC_rbr_inK54AicSCG :
STRUCT
	DTC: UDINT := 16#032C00;
	DFCid: UINT := 175;
	debounceMethod: USINT := TIME_UP_DOWN;
END_STRUCT
END_TYPE

(* ---- dfc_rbr_ink54or-DFC_rbr_inK54OR.st ---- *)
(* --- Interface --- *)
{attribute 'external_name' := 'cmp_rts_DFC_rbr_inK54OR'}
TYPE DFC_rbr_inK54OR :
STRUCT
	DTC: UDINT := 16#032D00;
	DFCid: UINT := 176;
	debounceMethod: USINT := TIME_UP_DOWN;
END_STRUCT
END_TYPE

(* ---- dfc_rbr_ink54scb-DFC_rbr_inK54SCB.st ---- *)
(* --- Interface --- *)
{attribute 'external_name' := 'cmp_rts_DFC_rbr_inK54SCB'}
TYPE DFC_rbr_inK54SCB :
STRUCT
	DTC: UDINT := 16#032E00;
	DFCid: UINT := 177;
	debounceMethod: USINT := TIME_UP_DOWN;
END_STRUCT
END_TYPE

(* ---- dfc_rbr_ink54scg-DFC_rbr_inK54SCG.st ---- *)
(* --- Interface --- *)
{attribute 'external_name' := 'cmp_rts_DFC_rbr_inK54SCG'}
TYPE DFC_rbr_inK54SCG :
STRUCT
	DTC: UDINT := 16#032F00;
	DFCid: UINT := 178;
	debounceMethod: USINT := TIME_UP_DOWN;
END_STRUCT
END_TYPE

(* ---- dfc_rbr_ink54shuntscb-DFC_rbr_inK54ShuntSCB.st ---- *)
(* --- Interface --- *)
{attribute 'external_name' := 'cmp_rts_DFC_rbr_inK54ShuntSCB'}
TYPE DFC_rbr_inK54ShuntSCB :
STRUCT
	DTC: UDINT := 16#033000;
	DFCid: UINT := 179;
	debounceMethod: USINT := TIME_UP_DOWN;
END_STRUCT
END_TYPE

(* ---- dfc_rbr_ink55aicscb-DFC_rbr_inK55AicSCB.st ---- *)
(* --- Interface --- *)
{attribute 'external_name' := 'cmp_rts_DFC_rbr_inK55AicSCB'}
TYPE DFC_rbr_inK55AicSCB :
STRUCT
	DTC: UDINT := 16#033100;
	DFCid: UINT := 180;
	debounceMethod: USINT := TIME_UP_DOWN;
END_STRUCT
END_TYPE

(* ---- dfc_rbr_ink55aicscg-DFC_rbr_inK55AicSCG.st ---- *)
(* --- Interface --- *)
{attribute 'external_name' := 'cmp_rts_DFC_rbr_inK55AicSCG'}
TYPE DFC_rbr_inK55AicSCG :
STRUCT
	DTC: UDINT := 16#033200;
	DFCid: UINT := 181;
	debounceMethod: USINT := TIME_UP_DOWN;
END_STRUCT
END_TYPE

(* ---- dfc_rbr_ink55or-DFC_rbr_inK55OR.st ---- *)
(* --- Interface --- *)
{attribute 'external_name' := 'cmp_rts_DFC_rbr_inK55OR'}
TYPE DFC_rbr_inK55OR :
STRUCT
	DTC: UDINT := 16#033300;
	DFCid: UINT := 182;
	debounceMethod: USINT := TIME_UP_DOWN;
END_STRUCT
END_TYPE

(* ---- dfc_rbr_ink55scb-DFC_rbr_inK55SCB.st ---- *)
(* --- Interface --- *)
{attribute 'external_name' := 'cmp_rts_DFC_rbr_inK55SCB'}
TYPE DFC_rbr_inK55SCB :
STRUCT
	DTC: UDINT := 16#033400;
	DFCid: UINT := 183;
	debounceMethod: USINT := TIME_UP_DOWN;
END_STRUCT
END_TYPE

(* ---- dfc_rbr_ink55scg-DFC_rbr_inK55SCG.st ---- *)
(* --- Interface --- *)
{attribute 'external_name' := 'cmp_rts_DFC_rbr_inK55SCG'}
TYPE DFC_rbr_inK55SCG :
STRUCT
	DTC: UDINT := 16#033500;
	DFCid: UINT := 184;
	debounceMethod: USINT := TIME_UP_DOWN;
END_STRUCT
END_TYPE

(* ---- dfc_rbr_ink55shuntscb-DFC_rbr_inK55ShuntSCB.st ---- *)
(* --- Interface --- *)
{attribute 'external_name' := 'cmp_rts_DFC_rbr_inK55ShuntSCB'}
TYPE DFC_rbr_inK55ShuntSCB :
STRUCT
	DTC: UDINT := 16#033600;
	DFCid: UINT := 185;
	debounceMethod: USINT := TIME_UP_DOWN;
END_STRUCT
END_TYPE

(* ---- dfc_rbr_ink56or-DFC_rbr_inK56OR.st ---- *)
(* --- Interface --- *)
{attribute 'external_name' := 'cmp_rts_DFC_rbr_inK56OR'}
TYPE DFC_rbr_inK56OR :
STRUCT
	DTC: UDINT := 16#033700;
	DFCid: UINT := 186;
	debounceMethod: USINT := TIME_UP_DOWN;
END_STRUCT
END_TYPE

(* ---- dfc_rbr_ink56scb-DFC_rbr_inK56SCB.st ---- *)
(* --- Interface --- *)
{attribute 'external_name' := 'cmp_rts_DFC_rbr_inK56SCB'}
TYPE DFC_rbr_inK56SCB :
STRUCT
	DTC: UDINT := 16#033800;
	DFCid: UINT := 187;
	debounceMethod: USINT := TIME_UP_DOWN;
END_STRUCT
END_TYPE

(* ---- dfc_rbr_ink56scg-DFC_rbr_inK56SCG.st ---- *)
(* --- Interface --- *)
{attribute 'external_name' := 'cmp_rts_DFC_rbr_inK56SCG'}
TYPE DFC_rbr_inK56SCG :
STRUCT
	DTC: UDINT := 16#033900;
	DFCid: UINT := 188;
	debounceMethod: USINT := TIME_UP_DOWN;
END_STRUCT
END_TYPE

(* ---- dfc_rbr_ink57or-DFC_rbr_inK57OR.st ---- *)
(* --- Interface --- *)
{attribute 'external_name' := 'cmp_rts_DFC_rbr_inK57OR'}
TYPE DFC_rbr_inK57OR :
STRUCT
	DTC: UDINT := 16#033A00;
	DFCid: UINT := 189;
	debounceMethod: USINT := TIME_UP_DOWN;
END_STRUCT
END_TYPE

(* ---- dfc_rbr_ink57scb-DFC_rbr_inK57SCB.st ---- *)
(* --- Interface --- *)
{attribute 'external_name' := 'cmp_rts_DFC_rbr_inK57SCB'}
TYPE DFC_rbr_inK57SCB :
STRUCT
	DTC: UDINT := 16#033B00;
	DFCid: UINT := 190;
	debounceMethod: USINT := TIME_UP_DOWN;
END_STRUCT
END_TYPE

(* ---- dfc_rbr_ink57scg-DFC_rbr_inK57SCG.st ---- *)
(* --- Interface --- *)
{attribute 'external_name' := 'cmp_rts_DFC_rbr_inK57SCG'}
TYPE DFC_rbr_inK57SCG :
STRUCT
	DTC: UDINT := 16#033C00;
	DFCid: UINT := 191;
	debounceMethod: USINT := TIME_UP_DOWN;
END_STRUCT
END_TYPE

(* ---- dfc_rbr_ink58or-DFC_rbr_inK58OR.st ---- *)
(* --- Interface --- *)
{attribute 'external_name' := 'cmp_rts_DFC_rbr_inK58OR'}
TYPE DFC_rbr_inK58OR :
STRUCT
	DTC: UDINT := 16#033D00;
	DFCid: UINT := 192;
	debounceMethod: USINT := TIME_UP_DOWN;
END_STRUCT
END_TYPE

(* ---- dfc_rbr_ink58scb-DFC_rbr_inK58SCB.st ---- *)
(* --- Interface --- *)
{attribute 'external_name' := 'cmp_rts_DFC_rbr_inK58SCB'}
TYPE DFC_rbr_inK58SCB :
STRUCT
	DTC: UDINT := 16#033E00;
	DFCid: UINT := 193;
	debounceMethod: USINT := TIME_UP_DOWN;
END_STRUCT
END_TYPE

(* ---- dfc_rbr_ink58scg-DFC_rbr_inK58SCG.st ---- *)
(* --- Interface --- *)
{attribute 'external_name' := 'cmp_rts_DFC_rbr_inK58SCG'}
TYPE DFC_rbr_inK58SCG :
STRUCT
	DTC: UDINT := 16#033F00;
	DFCid: UINT := 194;
	debounceMethod: USINT := TIME_UP_DOWN;
END_STRUCT
END_TYPE

(* ---- dfc_rbr_ink59or-DFC_rbr_inK59OR.st ---- *)
(* --- Interface --- *)
{attribute 'external_name' := 'cmp_rts_DFC_rbr_inK59OR'}
TYPE DFC_rbr_inK59OR :
STRUCT
	DTC: UDINT := 16#034000;
	DFCid: UINT := 195;
	debounceMethod: USINT := TIME_UP_DOWN;
END_STRUCT
END_TYPE

(* ---- dfc_rbr_ink59scb-DFC_rbr_inK59SCB.st ---- *)
(* --- Interface --- *)
{attribute 'external_name' := 'cmp_rts_DFC_rbr_inK59SCB'}
TYPE DFC_rbr_inK59SCB :
STRUCT
	DTC: UDINT := 16#034100;
	DFCid: UINT := 196;
	debounceMethod: USINT := TIME_UP_DOWN;
END_STRUCT
END_TYPE

(* ---- dfc_rbr_ink59scg-DFC_rbr_inK59SCG.st ---- *)
(* --- Interface --- *)
{attribute 'external_name' := 'cmp_rts_DFC_rbr_inK59SCG'}
TYPE DFC_rbr_inK59SCG :
STRUCT
	DTC: UDINT := 16#034200;
	DFCid: UINT := 197;
	debounceMethod: USINT := TIME_UP_DOWN;
END_STRUCT
END_TYPE

(* ---- dfc_rbr_ink60or-DFC_rbr_inK60OR.st ---- *)
(* --- Interface --- *)
{attribute 'external_name' := 'cmp_rts_DFC_rbr_inK60OR'}
TYPE DFC_rbr_inK60OR :
STRUCT
	DTC: UDINT := 16#034300;
	DFCid: UINT := 198;
	debounceMethod: USINT := TIME_UP_DOWN;
END_STRUCT
END_TYPE

(* ---- dfc_rbr_ink60scb-DFC_rbr_inK60SCB.st ---- *)
(* --- Interface --- *)
{attribute 'external_name' := 'cmp_rts_DFC_rbr_inK60SCB'}
TYPE DFC_rbr_inK60SCB :
STRUCT
	DTC: UDINT := 16#034400;
	DFCid: UINT := 199;
	debounceMethod: USINT := TIME_UP_DOWN;
END_STRUCT
END_TYPE

(* ---- dfc_rbr_ink60scg-DFC_rbr_inK60SCG.st ---- *)
(* --- Interface --- *)
{attribute 'external_name' := 'cmp_rts_DFC_rbr_inK60SCG'}
TYPE DFC_rbr_inK60SCG :
STRUCT
	DTC: UDINT := 16#034500;
	DFCid: UINT := 200;
	debounceMethod: USINT := TIME_UP_DOWN;
END_STRUCT
END_TYPE

(* ---- dfc_rbr_ink61aicscb-DFC_rbr_inK61AicSCB.st ---- *)
(* --- Interface --- *)
{attribute 'external_name' := 'cmp_rts_DFC_rbr_inK61AicSCB'}
TYPE DFC_rbr_inK61AicSCB :
STRUCT
	DTC: UDINT := 16#034600;
	DFCid: UINT := 201;
	debounceMethod: USINT := TIME_UP_DOWN;
END_STRUCT
END_TYPE

(* ---- dfc_rbr_ink61aicscg-DFC_rbr_inK61AicSCG.st ---- *)
(* --- Interface --- *)
{attribute 'external_name' := 'cmp_rts_DFC_rbr_inK61AicSCG'}
TYPE DFC_rbr_inK61AicSCG :
STRUCT
	DTC: UDINT := 16#034700;
	DFCid: UINT := 202;
	debounceMethod: USINT := TIME_UP_DOWN;
END_STRUCT
END_TYPE

(* ---- dfc_rbr_ink61or-DFC_rbr_inK61OR.st ---- *)
(* --- Interface --- *)
{attribute 'external_name' := 'cmp_rts_DFC_rbr_inK61OR'}
TYPE DFC_rbr_inK61OR :
STRUCT
	DTC: UDINT := 16#034800;
	DFCid: UINT := 203;
	debounceMethod: USINT := TIME_UP_DOWN;
END_STRUCT
END_TYPE

(* ---- dfc_rbr_ink61scb-DFC_rbr_inK61SCB.st ---- *)
(* --- Interface --- *)
{attribute 'external_name' := 'cmp_rts_DFC_rbr_inK61SCB'}
TYPE DFC_rbr_inK61SCB :
STRUCT
	DTC: UDINT := 16#034900;
	DFCid: UINT := 204;
	debounceMethod: USINT := TIME_UP_DOWN;
END_STRUCT
END_TYPE

(* ---- dfc_rbr_ink61scg-DFC_rbr_inK61SCG.st ---- *)
(* --- Interface --- *)
{attribute 'external_name' := 'cmp_rts_DFC_rbr_inK61SCG'}
TYPE DFC_rbr_inK61SCG :
STRUCT
	DTC: UDINT := 16#034A00;
	DFCid: UINT := 205;
	debounceMethod: USINT := TIME_UP_DOWN;
END_STRUCT
END_TYPE

(* ---- dfc_rbr_ink61shuntscb-DFC_rbr_inK61ShuntSCB.st ---- *)
(* --- Interface --- *)
{attribute 'external_name' := 'cmp_rts_DFC_rbr_inK61ShuntSCB'}
TYPE DFC_rbr_inK61ShuntSCB :
STRUCT
	DTC: UDINT := 16#034B00;
	DFCid: UINT := 206;
	debounceMethod: USINT := TIME_UP_DOWN;
END_STRUCT
END_TYPE

(* ---- dfc_rbr_ink62or-DFC_rbr_inK62OR.st ---- *)
(* --- Interface --- *)
{attribute 'external_name' := 'cmp_rts_DFC_rbr_inK62OR'}
TYPE DFC_rbr_inK62OR :
STRUCT
	DTC: UDINT := 16#034C00;
	DFCid: UINT := 207;
	debounceMethod: USINT := TIME_UP_DOWN;
END_STRUCT
END_TYPE

(* ---- dfc_rbr_ink62scb-DFC_rbr_inK62SCB.st ---- *)
(* --- Interface --- *)
{attribute 'external_name' := 'cmp_rts_DFC_rbr_inK62SCB'}
TYPE DFC_rbr_inK62SCB :
STRUCT
	DTC: UDINT := 16#034D00;
	DFCid: UINT := 208;
	debounceMethod: USINT := TIME_UP_DOWN;
END_STRUCT
END_TYPE

(* ---- dfc_rbr_ink62scg-DFC_rbr_inK62SCG.st ---- *)
(* --- Interface --- *)
{attribute 'external_name' := 'cmp_rts_DFC_rbr_inK62SCG'}
TYPE DFC_rbr_inK62SCG :
STRUCT
	DTC: UDINT := 16#034E00;
	DFCid: UINT := 209;
	debounceMethod: USINT := TIME_UP_DOWN;
END_STRUCT
END_TYPE

(* ---- dfc_rbr_ink63aicscb-DFC_rbr_inK63AicSCB.st ---- *)
(* --- Interface --- *)
{attribute 'external_name' := 'cmp_rts_DFC_rbr_inK63AicSCB'}
TYPE DFC_rbr_inK63AicSCB :
STRUCT
	DTC: UDINT := 16#03CF00;
	DFCid: UINT := 210;
	debounceMethod: USINT := TIME_UP_DOWN;
END_STRUCT
END_TYPE

(* ---- dfc_rbr_ink63aicscg-DFC_rbr_inK63AicSCG.st ---- *)
(* --- Interface --- *)
{attribute 'external_name' := 'cmp_rts_DFC_rbr_inK63AicSCG'}
TYPE DFC_rbr_inK63AicSCG :
STRUCT
	DTC: UDINT := 16#03D000;
	DFCid: UINT := 211;
	debounceMethod: USINT := TIME_UP_DOWN;
END_STRUCT
END_TYPE

(* ---- dfc_rbr_ink63or-DFC_rbr_inK63OR.st ---- *)
(* --- Interface --- *)
{attribute 'external_name' := 'cmp_rts_DFC_rbr_inK63OR'}
TYPE DFC_rbr_inK63OR :
STRUCT
	DTC: UDINT := 16#034F00;
	DFCid: UINT := 212;
	debounceMethod: USINT := TIME_UP_DOWN;
END_STRUCT
END_TYPE

(* ---- dfc_rbr_ink63scb-DFC_rbr_inK63SCB.st ---- *)
(* --- Interface --- *)
{attribute 'external_name' := 'cmp_rts_DFC_rbr_inK63SCB'}
TYPE DFC_rbr_inK63SCB :
STRUCT
	DTC: UDINT := 16#035000;
	DFCid: UINT := 213;
	debounceMethod: USINT := TIME_UP_DOWN;
END_STRUCT
END_TYPE

(* ---- dfc_rbr_ink63scg-DFC_rbr_inK63SCG.st ---- *)
(* --- Interface --- *)
{attribute 'external_name' := 'cmp_rts_DFC_rbr_inK63SCG'}
TYPE DFC_rbr_inK63SCG :
STRUCT
	DTC: UDINT := 16#035100;
	DFCid: UINT := 214;
	debounceMethod: USINT := TIME_UP_DOWN;
END_STRUCT
END_TYPE

(* ---- dfc_rbr_ink63shuntscb-DFC_rbr_inK63ShuntSCB.st ---- *)
(* --- Interface --- *)
{attribute 'external_name' := 'cmp_rts_DFC_rbr_inK63ShuntSCB'}
TYPE DFC_rbr_inK63ShuntSCB :
STRUCT
	DTC: UDINT := 16#03D100;
	DFCid: UINT := 215;
	debounceMethod: USINT := TIME_UP_DOWN;
END_STRUCT
END_TYPE

(* ---- dfc_rbr_ink64aicscb-DFC_rbr_inK64AicSCB.st ---- *)
(* --- Interface --- *)
{attribute 'external_name' := 'cmp_rts_DFC_rbr_inK64AicSCB'}
TYPE DFC_rbr_inK64AicSCB :
STRUCT
	DTC: UDINT := 16#03D200;
	DFCid: UINT := 216;
	debounceMethod: USINT := TIME_UP_DOWN;
END_STRUCT
END_TYPE

(* ---- dfc_rbr_ink64aicscg-DFC_rbr_inK64AicSCG.st ---- *)
(* --- Interface --- *)
{attribute 'external_name' := 'cmp_rts_DFC_rbr_inK64AicSCG'}
TYPE DFC_rbr_inK64AicSCG :
STRUCT
	DTC: UDINT := 16#03D300;
	DFCid: UINT := 217;
	debounceMethod: USINT := TIME_UP_DOWN;
END_STRUCT
END_TYPE

(* ---- dfc_rbr_ink64or-DFC_rbr_inK64OR.st ---- *)
(* --- Interface --- *)
{attribute 'external_name' := 'cmp_rts_DFC_rbr_inK64OR'}
TYPE DFC_rbr_inK64OR :
STRUCT
	DTC: UDINT := 16#035200;
	DFCid: UINT := 218;
	debounceMethod: USINT := TIME_UP_DOWN;
END_STRUCT
END_TYPE

(* ---- dfc_rbr_ink64scb-DFC_rbr_inK64SCB.st ---- *)
(* --- Interface --- *)
{attribute 'external_name' := 'cmp_rts_DFC_rbr_inK64SCB'}
TYPE DFC_rbr_inK64SCB :
STRUCT
	DTC: UDINT := 16#035300;
	DFCid: UINT := 219;
	debounceMethod: USINT := TIME_UP_DOWN;
END_STRUCT
END_TYPE

(* ---- dfc_rbr_ink64scg-DFC_rbr_inK64SCG.st ---- *)
(* --- Interface --- *)
{attribute 'external_name' := 'cmp_rts_DFC_rbr_inK64SCG'}
TYPE DFC_rbr_inK64SCG :
STRUCT
	DTC: UDINT := 16#035400;
	DFCid: UINT := 220;
	debounceMethod: USINT := TIME_UP_DOWN;
END_STRUCT
END_TYPE

(* ---- dfc_rbr_ink64shuntscb-DFC_rbr_inK64ShuntSCB.st ---- *)
(* --- Interface --- *)
{attribute 'external_name' := 'cmp_rts_DFC_rbr_inK64ShuntSCB'}
TYPE DFC_rbr_inK64ShuntSCB :
STRUCT
	DTC: UDINT := 16#03D400;
	DFCid: UINT := 221;
	debounceMethod: USINT := TIME_UP_DOWN;
END_STRUCT
END_TYPE

(* ---- dfc_rbr_ink65aicscb-DFC_rbr_inK65AicSCB.st ---- *)
(* --- Interface --- *)
{attribute 'external_name' := 'cmp_rts_DFC_rbr_inK65AicSCB'}
TYPE DFC_rbr_inK65AicSCB :
STRUCT
	DTC: UDINT := 16#03D500;
	DFCid: UINT := 222;
	debounceMethod: USINT := TIME_UP_DOWN;
END_STRUCT
END_TYPE

(* ---- dfc_rbr_ink65aicscg-DFC_rbr_inK65AicSCG.st ---- *)
(* --- Interface --- *)
{attribute 'external_name' := 'cmp_rts_DFC_rbr_inK65AicSCG'}
TYPE DFC_rbr_inK65AicSCG :
STRUCT
	DTC: UDINT := 16#03D600;
	DFCid: UINT := 223;
	debounceMethod: USINT := TIME_UP_DOWN;
END_STRUCT
END_TYPE

(* ---- dfc_rbr_ink65or-DFC_rbr_inK65OR.st ---- *)
(* --- Interface --- *)
{attribute 'external_name' := 'cmp_rts_DFC_rbr_inK65OR'}
TYPE DFC_rbr_inK65OR :
STRUCT
	DTC: UDINT := 16#035500;
	DFCid: UINT := 224;
	debounceMethod: USINT := TIME_UP_DOWN;
END_STRUCT
END_TYPE

(* ---- dfc_rbr_ink65scb-DFC_rbr_inK65SCB.st ---- *)
(* --- Interface --- *)
{attribute 'external_name' := 'cmp_rts_DFC_rbr_inK65SCB'}
TYPE DFC_rbr_inK65SCB :
STRUCT
	DTC: UDINT := 16#035600;
	DFCid: UINT := 225;
	debounceMethod: USINT := TIME_UP_DOWN;
END_STRUCT
END_TYPE

(* ---- dfc_rbr_ink65scg-DFC_rbr_inK65SCG.st ---- *)
(* --- Interface --- *)
{attribute 'external_name' := 'cmp_rts_DFC_rbr_inK65SCG'}
TYPE DFC_rbr_inK65SCG :
STRUCT
	DTC: UDINT := 16#035700;
	DFCid: UINT := 226;
	debounceMethod: USINT := TIME_UP_DOWN;
END_STRUCT
END_TYPE

(* ---- dfc_rbr_ink65shuntscb-DFC_rbr_inK65ShuntSCB.st ---- *)
(* --- Interface --- *)
{attribute 'external_name' := 'cmp_rts_DFC_rbr_inK65ShuntSCB'}
TYPE DFC_rbr_inK65ShuntSCB :
STRUCT
	DTC: UDINT := 16#03D700;
	DFCid: UINT := 227;
	debounceMethod: USINT := TIME_UP_DOWN;
END_STRUCT
END_TYPE

(* ---- dfc_rbr_ink74or-DFC_rbr_inK74OR.st ---- *)
(* --- Interface --- *)
{attribute 'external_name' := 'cmp_rts_DFC_rbr_inK74OR'}
TYPE DFC_rbr_inK74OR :
STRUCT
	DTC: UDINT := 16#035800;
	DFCid: UINT := 228;
	debounceMethod: USINT := TIME_UP_DOWN;
END_STRUCT
END_TYPE

(* ---- dfc_rbr_ink74scb-DFC_rbr_inK74SCB.st ---- *)
(* --- Interface --- *)
{attribute 'external_name' := 'cmp_rts_DFC_rbr_inK74SCB'}
TYPE DFC_rbr_inK74SCB :
STRUCT
	DTC: UDINT := 16#035900;
	DFCid: UINT := 229;
	debounceMethod: USINT := TIME_UP_DOWN;
END_STRUCT
END_TYPE

(* ---- dfc_rbr_ink74scg-DFC_rbr_inK74SCG.st ---- *)
(* --- Interface --- *)
{attribute 'external_name' := 'cmp_rts_DFC_rbr_inK74SCG'}
TYPE DFC_rbr_inK74SCG :
STRUCT
	DTC: UDINT := 16#035A00;
	DFCid: UINT := 230;
	debounceMethod: USINT := TIME_UP_DOWN;
END_STRUCT
END_TYPE

(* ---- dfc_rbr_ink75or-DFC_rbr_inK75OR.st ---- *)
(* --- Interface --- *)
{attribute 'external_name' := 'cmp_rts_DFC_rbr_inK75OR'}
TYPE DFC_rbr_inK75OR :
STRUCT
	DTC: UDINT := 16#035B00;
	DFCid: UINT := 231;
	debounceMethod: USINT := TIME_UP_DOWN;
END_STRUCT
END_TYPE

(* ---- dfc_rbr_ink75scb-DFC_rbr_inK75SCB.st ---- *)
(* --- Interface --- *)
{attribute 'external_name' := 'cmp_rts_DFC_rbr_inK75SCB'}
TYPE DFC_rbr_inK75SCB :
STRUCT
	DTC: UDINT := 16#035C00;
	DFCid: UINT := 232;
	debounceMethod: USINT := TIME_UP_DOWN;
END_STRUCT
END_TYPE

(* ---- dfc_rbr_ink75scg-DFC_rbr_inK75SCG.st ---- *)
(* --- Interface --- *)
{attribute 'external_name' := 'cmp_rts_DFC_rbr_inK75SCG'}
TYPE DFC_rbr_inK75SCG :
STRUCT
	DTC: UDINT := 16#035D00;
	DFCid: UINT := 233;
	debounceMethod: USINT := TIME_UP_DOWN;
END_STRUCT
END_TYPE

(* ---- dfc_rbr_ink76or-DFC_rbr_inK76OR.st ---- *)
(* --- Interface --- *)
{attribute 'external_name' := 'cmp_rts_DFC_rbr_inK76OR'}
TYPE DFC_rbr_inK76OR :
STRUCT
	DTC: UDINT := 16#035E00;
	DFCid: UINT := 234;
	debounceMethod: USINT := TIME_UP_DOWN;
END_STRUCT
END_TYPE

(* ---- dfc_rbr_ink76scb-DFC_rbr_inK76SCB.st ---- *)
(* --- Interface --- *)
{attribute 'external_name' := 'cmp_rts_DFC_rbr_inK76SCB'}
TYPE DFC_rbr_inK76SCB :
STRUCT
	DTC: UDINT := 16#035F00;
	DFCid: UINT := 235;
	debounceMethod: USINT := TIME_UP_DOWN;
END_STRUCT
END_TYPE

(* ---- dfc_rbr_ink76scg-DFC_rbr_inK76SCG.st ---- *)
(* --- Interface --- *)
{attribute 'external_name' := 'cmp_rts_DFC_rbr_inK76SCG'}
TYPE DFC_rbr_inK76SCG :
STRUCT
	DTC: UDINT := 16#036000;
	DFCid: UINT := 236;
	debounceMethod: USINT := TIME_UP_DOWN;
END_STRUCT
END_TYPE

(* ---- dfc_rbr_ink77or-DFC_rbr_inK77OR.st ---- *)
(* --- Interface --- *)
{attribute 'external_name' := 'cmp_rts_DFC_rbr_inK77OR'}
TYPE DFC_rbr_inK77OR :
STRUCT
	DTC: UDINT := 16#036100;
	DFCid: UINT := 237;
	debounceMethod: USINT := TIME_UP_DOWN;
END_STRUCT
END_TYPE

(* ---- dfc_rbr_ink77scb-DFC_rbr_inK77SCB.st ---- *)
(* --- Interface --- *)
{attribute 'external_name' := 'cmp_rts_DFC_rbr_inK77SCB'}
TYPE DFC_rbr_inK77SCB :
STRUCT
	DTC: UDINT := 16#036200;
	DFCid: UINT := 238;
	debounceMethod: USINT := TIME_UP_DOWN;
END_STRUCT
END_TYPE

(* ---- dfc_rbr_ink77scg-DFC_rbr_inK77SCG.st ---- *)
(* --- Interface --- *)
{attribute 'external_name' := 'cmp_rts_DFC_rbr_inK77SCG'}
TYPE DFC_rbr_inK77SCG :
STRUCT
	DTC: UDINT := 16#036300;
	DFCid: UINT := 239;
	debounceMethod: USINT := TIME_UP_DOWN;
END_STRUCT
END_TYPE

(* ---- dfc_rbr_ink78or-DFC_rbr_inK78OR.st ---- *)
(* --- Interface --- *)
{attribute 'external_name' := 'cmp_rts_DFC_rbr_inK78OR'}
TYPE DFC_rbr_inK78OR :
STRUCT
	DTC: UDINT := 16#036400;
	DFCid: UINT := 240;
	debounceMethod: USINT := TIME_UP_DOWN;
END_STRUCT
END_TYPE

(* ---- dfc_rbr_ink78scb-DFC_rbr_inK78SCB.st ---- *)
(* --- Interface --- *)
{attribute 'external_name' := 'cmp_rts_DFC_rbr_inK78SCB'}
TYPE DFC_rbr_inK78SCB :
STRUCT
	DTC: UDINT := 16#036500;
	DFCid: UINT := 241;
	debounceMethod: USINT := TIME_UP_DOWN;
END_STRUCT
END_TYPE

(* ---- dfc_rbr_ink78scg-DFC_rbr_inK78SCG.st ---- *)
(* --- Interface --- *)
{attribute 'external_name' := 'cmp_rts_DFC_rbr_inK78SCG'}
TYPE DFC_rbr_inK78SCG :
STRUCT
	DTC: UDINT := 16#036600;
	DFCid: UINT := 242;
	debounceMethod: USINT := TIME_UP_DOWN;
END_STRUCT
END_TYPE

(* ---- dfc_rbr_inphase-DFC_rbr_inPhase.st ---- *)
(* --- Interface --- *)
{attribute 'external_name' := 'cmp_rts_DFC_rbr_inPhase'}
TYPE DFC_rbr_inPhase :
STRUCT
	DTC: UDINT := 16#039E00;
	DFCid: UINT := 592;
	debounceMethod: USINT := NO_DEBOUNCE;
END_STRUCT
END_TYPE

(* ---- dfc_rbr_inphasegetstatus-DFC_rbr_inPhaseGetStatus.st ---- *)
(* --- Interface --- *)
{attribute 'external_name' := 'cmp_rts_DFC_rbr_inPhaseGetStatus'}
TYPE DFC_rbr_inPhaseGetStatus :
STRUCT
	DTC: UDINT := 16#039F00;
	DFCid: UINT := 593;
	debounceMethod: USINT := NO_DEBOUNCE;
END_STRUCT
END_TYPE

(* ---- dfc_rbr_inphaseresetcounter-DFC_rbr_inPhaseResetCounter.st ---- *)
(* --- Interface --- *)
{attribute 'external_name' := 'cmp_rts_DFC_rbr_inPhaseResetCounter'}
TYPE DFC_rbr_inPhaseResetCounter :
STRUCT
	DTC: UDINT := 16#03A000;
	DFCid: UINT := 594;
	debounceMethod: USINT := NO_DEBOUNCE;
END_STRUCT
END_TYPE

(* ---- dfc_rbr_inri-DFC_rbr_inRi.st ---- *)
(* --- Interface --- *)
{attribute 'external_name' := 'cmp_rts_DFC_rbr_inRi'}
TYPE DFC_rbr_inRi :
STRUCT
	DTC: UDINT := 16#038A00;
	DFCid: UINT := 595;
	debounceMethod: USINT := NO_DEBOUNCE;
END_STRUCT
END_TYPE

(* ---- dfc_rbr_inricfg-DFC_rbr_inRiCfg.st ---- *)
(* --- Interface --- *)
{attribute 'external_name' := 'cmp_rts_DFC_rbr_inRiCfg'}
TYPE DFC_rbr_inRiCfg :
STRUCT
	DTC: UDINT := 16#038B00;
	DFCid: UINT := 596;
	debounceMethod: USINT := NO_DEBOUNCE;
END_STRUCT
END_TYPE

(* ---- dfc_rbr_inricfgtemp-DFC_rbr_inRiCfgTemp.st ---- *)
(* --- Interface --- *)
{attribute 'external_name' := 'cmp_rts_DFC_rbr_inRiCfgTemp'}
TYPE DFC_rbr_inRiCfgTemp :
STRUCT
	DTC: UDINT := 16#039C00;
	DFCid: UINT := 597;
	debounceMethod: USINT := NO_DEBOUNCE;
END_STRUCT
END_TYPE

(* ---- dfc_rbr_inrigetstatus-DFC_rbr_inRiGetStatus.st ---- *)
(* --- Interface --- *)
{attribute 'external_name' := 'cmp_rts_DFC_rbr_inRiGetStatus'}
TYPE DFC_rbr_inRiGetStatus :
STRUCT
	DTC: UDINT := 16#038E00;
	DFCid: UINT := 598;
	debounceMethod: USINT := NO_DEBOUNCE;
END_STRUCT
END_TYPE

(* ---- dfc_rbr_inrigettemp-DFC_rbr_inRiGetTemp.st ---- *)
(* --- Interface --- *)
{attribute 'external_name' := 'cmp_rts_DFC_rbr_inRiGetTemp'}
TYPE DFC_rbr_inRiGetTemp :
STRUCT
	DTC: UDINT := 16#039D00;
	DFCid: UINT := 599;
	debounceMethod: USINT := NO_DEBOUNCE;
END_STRUCT
END_TYPE

(* ---- dfc_rbr_insentcopyfdfifo-DFC_rbr_inSentCopyFDFifo.st ---- *)
(* --- Interface --- *)
{attribute 'external_name' := 'cmp_rts_DFC_rbr_inSentCopyFDFifo'}
TYPE DFC_rbr_inSentCopyFDFifo :
STRUCT
	DTC: UDINT := 16#039800;
	DFCid: UINT := 600;
	debounceMethod: USINT := NO_DEBOUNCE;
END_STRUCT
END_TYPE

(* ---- dfc_rbr_insentdisable-DFC_rbr_inSentDisable.st ---- *)
(* --- Interface --- *)
{attribute 'external_name' := 'cmp_rts_DFC_rbr_inSentDisable'}
TYPE DFC_rbr_inSentDisable :
STRUCT
	DTC: UDINT := 16#039100;
	DFCid: UINT := 601;
	debounceMethod: USINT := NO_DEBOUNCE;
END_STRUCT
END_TYPE

(* ---- dfc_rbr_insentenable-DFC_rbr_inSentEnable.st ---- *)
(* --- Interface --- *)
{attribute 'external_name' := 'cmp_rts_DFC_rbr_inSentEnable'}
TYPE DFC_rbr_inSentEnable :
STRUCT
	DTC: UDINT := 16#039000;
	DFCid: UINT := 602;
	debounceMethod: USINT := NO_DEBOUNCE;
END_STRUCT
END_TYPE

(* ---- dfc_rbr_insentgeterrorstatus-DFC_rbr_inSentGetErrorStatus.st ---- *)
(* --- Interface --- *)
{attribute 'external_name' := 'cmp_rts_DFC_rbr_inSentGetErrorStatus'}
TYPE DFC_rbr_inSentGetErrorStatus :
STRUCT
	DTC: UDINT := 16#039500;
	DFCid: UINT := 603;
	debounceMethod: USINT := NO_DEBOUNCE;
END_STRUCT
END_TYPE

(* ---- dfc_rbr_insentgetfd-DFC_rbr_inSentGetFD.st ---- *)
(* --- Interface --- *)
{attribute 'external_name' := 'cmp_rts_DFC_rbr_inSentGetFD'}
TYPE DFC_rbr_inSentGetFD :
STRUCT
	DTC: UDINT := 16#039200;
	DFCid: UINT := 604;
	debounceMethod: USINT := NO_DEBOUNCE;
END_STRUCT
END_TYPE

(* ---- dfc_rbr_insentgetsd-DFC_rbr_inSentGetSD.st ---- *)
(* --- Interface --- *)
{attribute 'external_name' := 'cmp_rts_DFC_rbr_inSentGetSD'}
TYPE DFC_rbr_inSentGetSD :
STRUCT
	DTC: UDINT := 16#039300;
	DFCid: UINT := 605;
	debounceMethod: USINT := NO_DEBOUNCE;
END_STRUCT
END_TYPE

(* ---- dfc_rbr_insentgetsddatabox-DFC_rbr_inSentGetSDDatabox.st ---- *)
(* --- Interface --- *)
{attribute 'external_name' := 'cmp_rts_DFC_rbr_inSentGetSDDatabox'}
TYPE DFC_rbr_inSentGetSDDatabox :
STRUCT
	DTC: UDINT := 16#039B00;
	DFCid: UINT := 606;
	debounceMethod: USINT := NO_DEBOUNCE;
END_STRUCT
END_TYPE

(* ---- dfc_rbr_insentgetstatus-DFC_rbr_inSentGetStatus.st ---- *)
(* --- Interface --- *)
{attribute 'external_name' := 'cmp_rts_DFC_rbr_inSentGetStatus'}
TYPE DFC_rbr_inSentGetStatus :
STRUCT
	DTC: UDINT := 16#039400;
	DFCid: UINT := 607;
	debounceMethod: USINT := NO_DEBOUNCE;
END_STRUCT
END_TYPE

(* ---- dfc_rbr_insentinitsddatabox-DFC_rbr_inSentInitSDDatabox.st ---- *)
(* --- Interface --- *)
{attribute 'external_name' := 'cmp_rts_DFC_rbr_inSentInitSDDatabox'}
TYPE DFC_rbr_inSentInitSDDatabox :
STRUCT
	DTC: UDINT := 16#039A00;
	DFCid: UINT := 608;
	debounceMethod: USINT := NO_DEBOUNCE;
END_STRUCT
END_TYPE

(* ---- dfc_rbr_insentregistercopyfdfifo-DFC_rbr_inSentRegisterCopyFDFifo.st ---- *)
(* --- Interface --- *)
{attribute 'external_name' := 'cmp_rts_DFC_rbr_inSentRegisterCopyFDFifo'}
TYPE DFC_rbr_inSentRegisterCopyFDFifo :
STRUCT
	DTC: UDINT := 16#039700;
	DFCid: UINT := 609;
	debounceMethod: USINT := NO_DEBOUNCE;
END_STRUCT
END_TYPE

(* ---- dfc_rbr_insentregisterfdfifo-DFC_rbr_inSentRegisterFDFifo.st ---- *)
(* --- Interface --- *)
{attribute 'external_name' := 'cmp_rts_DFC_rbr_inSentRegisterFDFifo'}
TYPE DFC_rbr_inSentRegisterFDFifo :
STRUCT
	DTC: UDINT := 16#039600;
	DFCid: UINT := 610;
	debounceMethod: USINT := NO_DEBOUNCE;
END_STRUCT
END_TYPE

(* ---- dfc_rbr_insentregistersddataboxes-DFC_rbr_inSentRegisterSDDataboxes.st ---- *)
(* --- Interface --- *)
{attribute 'external_name' := 'cmp_rts_DFC_rbr_inSentRegisterSDDataboxes'}
TYPE DFC_rbr_inSentRegisterSDDataboxes :
STRUCT
	DTC: UDINT := 16#039900;
	DFCid: UINT := 611;
	debounceMethod: USINT := NO_DEBOUNCE;
END_STRUCT
END_TYPE

(* ---- dfc_rbr_isobuscanrxbufferoverflow-DFC_rbr_isobusCanRxBufferOverflow.st ---- *)
(* --- Interface --- *)
{attribute 'external_name' := 'cmp_rts_DFC_rbr_isobusCanRxBufferOverflow'}
TYPE DFC_rbr_isobusCanRxBufferOverflow :
STRUCT
	DTC: UDINT := 16#050100;
	DFCid: UINT := 612;
	debounceMethod: USINT := NO_DEBOUNCE;
END_STRUCT
END_TYPE

(* ---- dfc_rbr_isobusgetcaaddrparam-DFC_rbr_isobusGetCaAddrParam.st ---- *)
(* --- Interface --- *)
{attribute 'external_name' := 'cmp_rts_DFC_rbr_isobusGetCaAddrParam'}
TYPE DFC_rbr_isobusGetCaAddrParam :
STRUCT
	DTC: UDINT := 16#050200;
	DFCid: UINT := 613;
	debounceMethod: USINT := NO_DEBOUNCE;
END_STRUCT
END_TYPE

(* ---- dfc_rbr_isobusgetdiagnosticparam-DFC_rbr_isobusGetDiagnosticParam.st ---- *)
(* --- Interface --- *)
{attribute 'external_name' := 'cmp_rts_DFC_rbr_isobusGetDiagnosticParam'}
TYPE DFC_rbr_isobusGetDiagnosticParam :
STRUCT
	DTC: UDINT := 16#050300;
	DFCid: UINT := 614;
	debounceMethod: USINT := NO_DEBOUNCE;
END_STRUCT
END_TYPE

(* ---- dfc_rbr_isobusgetrxdataboxstatusparam-DFC_rbr_isobusGetRxDataboxStatusParam.st ---- *)
(* --- Interface --- *)
{attribute 'external_name' := 'cmp_rts_DFC_rbr_isobusGetRxDataboxStatusParam'}
TYPE DFC_rbr_isobusGetRxDataboxStatusParam :
STRUCT
	DTC: UDINT := 16#050400;
	DFCid: UINT := 615;
	debounceMethod: USINT := NO_DEBOUNCE;
END_STRUCT
END_TYPE

(* ---- dfc_rbr_isobusgetstatusparam-DFC_rbr_isobusGetStatusParam.st ---- *)
(* --- Interface --- *)
{attribute 'external_name' := 'cmp_rts_DFC_rbr_isobusGetStatusParam'}
TYPE DFC_rbr_isobusGetStatusParam :
STRUCT
	DTC: UDINT := 16#050500;
	DFCid: UINT := 616;
	debounceMethod: USINT := NO_DEBOUNCE;
END_STRUCT
END_TYPE

(* ---- dfc_rbr_isobusinitcommcamissing-DFC_rbr_isobusInitCommCaMissing.st ---- *)
(* --- Interface --- *)
{attribute 'external_name' := 'cmp_rts_DFC_rbr_isobusInitCommCaMissing'}
TYPE DFC_rbr_isobusInitCommCaMissing :
STRUCT
	DTC: UDINT := 16#050600;
	DFCid: UINT := 617;
	debounceMethod: USINT := NO_DEBOUNCE;
END_STRUCT
END_TYPE

(* ---- dfc_rbr_isobusinitcommparam-DFC_rbr_isobusInitCommParam.st ---- *)
(* --- Interface --- *)
{attribute 'external_name' := 'cmp_rts_DFC_rbr_isobusInitCommParam'}
TYPE DFC_rbr_isobusInitCommParam :
STRUCT
	DTC: UDINT := 16#050700;
	DFCid: UINT := 618;
	debounceMethod: USINT := NO_DEBOUNCE;
END_STRUCT
END_TYPE

(* ---- dfc_rbr_isobusinitcommstate-DFC_rbr_isobusInitCommState.st ---- *)
(* --- Interface --- *)
{attribute 'external_name' := 'cmp_rts_DFC_rbr_isobusInitCommState'}
TYPE DFC_rbr_isobusInitCommState :
STRUCT
	DTC: UDINT := 16#050800;
	DFCid: UINT := 619;
	debounceMethod: USINT := NO_DEBOUNCE;
END_STRUCT
END_TYPE

(* ---- dfc_rbr_isobusinitdiagnosticparam-DFC_rbr_isobusInitDiagnosticParam.st ---- *)
(* --- Interface --- *)
{attribute 'external_name' := 'cmp_rts_DFC_rbr_isobusInitDiagnosticParam'}
TYPE DFC_rbr_isobusInitDiagnosticParam :
STRUCT
	DTC: UDINT := 16#050900;
	DFCid: UINT := 620;
	debounceMethod: USINT := NO_DEBOUNCE;
END_STRUCT
END_TYPE

(* ---- dfc_rbr_isobusinitfailurelistparam-DFC_rbr_isobusInitFailureListParam.st ---- *)
(* --- Interface --- *)
{attribute 'external_name' := 'cmp_rts_DFC_rbr_isobusInitFailureListParam'}
TYPE DFC_rbr_isobusInitFailureListParam :
STRUCT
	DTC: UDINT := 16#050A00;
	DFCid: UINT := 621;
	debounceMethod: USINT := NO_DEBOUNCE;
END_STRUCT
END_TYPE

(* ---- dfc_rbr_isobusinitrxdataboxparam-DFC_rbr_isobusInitRxDataboxParam.st ---- *)
(* --- Interface --- *)
{attribute 'external_name' := 'cmp_rts_DFC_rbr_isobusInitRxDataboxParam'}
TYPE DFC_rbr_isobusInitRxDataboxParam :
STRUCT
	DTC: UDINT := 16#050B00;
	DFCid: UINT := 622;
	debounceMethod: USINT := NO_DEBOUNCE;
END_STRUCT
END_TYPE

(* ---- dfc_rbr_isobusinittxdataboxparam-DFC_rbr_isobusInitTxDataboxParam.st ---- *)
(* --- Interface --- *)
{attribute 'external_name' := 'cmp_rts_DFC_rbr_isobusInitTxDataboxParam'}
TYPE DFC_rbr_isobusInitTxDataboxParam :
STRUCT
	DTC: UDINT := 16#050C00;
	DFCid: UINT := 623;
	debounceMethod: USINT := NO_DEBOUNCE;
END_STRUCT
END_TYPE

(* ---- dfc_rbr_isobusregistererrclrcallbackparam-DFC_rbr_isobusRegisterErrClrCallbackParam.st ---- *)
(* --- Interface --- *)
{attribute 'external_name' := 'cmp_rts_DFC_rbr_isobusRegisterErrClrCallbackParam'}
TYPE DFC_rbr_isobusRegisterErrClrCallbackParam :
STRUCT
	DTC: UDINT := 16#050D00;
	DFCid: UINT := 630;
	debounceMethod: USINT := NO_DEBOUNCE;
END_STRUCT
END_TYPE

(* ---- dfc_rbr_isobusregisterinstancesoverlap-DFC_rbr_isobusRegisterInstancesOverlap.st ---- *)
(* --- Interface --- *)
{attribute 'external_name' := 'cmp_rts_DFC_rbr_isobusRegisterInstancesOverlap'}
TYPE DFC_rbr_isobusRegisterInstancesOverlap :
STRUCT
	DTC: UDINT := 16#050E00;
	DFCid: UINT := 631;
	debounceMethod: USINT := NO_DEBOUNCE;
END_STRUCT
END_TYPE

(* ---- dfc_rbr_isobusregisterinstancesparam-DFC_rbr_isobusRegisterInstancesParam.st ---- *)
(* --- Interface --- *)
{attribute 'external_name' := 'cmp_rts_DFC_rbr_isobusRegisterInstancesParam'}
TYPE DFC_rbr_isobusRegisterInstancesParam :
STRUCT
	DTC: UDINT := 16#050F00;
	DFCid: UINT := 632;
	debounceMethod: USINT := NO_DEBOUNCE;
END_STRUCT
END_TYPE

(* ---- dfc_rbr_isobusregisterinstancesstate-DFC_rbr_isobusRegisterInstancesState.st ---- *)
(* --- Interface --- *)
{attribute 'external_name' := 'cmp_rts_DFC_rbr_isobusRegisterInstancesState'}
TYPE DFC_rbr_isobusRegisterInstancesState :
STRUCT
	DTC: UDINT := 16#051000;
	DFCid: UINT := 633;
	debounceMethod: USINT := NO_DEBOUNCE;
END_STRUCT
END_TYPE

(* ---- dfc_rbr_isobusregrxdataboxoverlap-DFC_rbr_isobusRegRxDataboxOverlap.st ---- *)
(* --- Interface --- *)
{attribute 'external_name' := 'cmp_rts_DFC_rbr_isobusRegRxDataboxOverlap'}
TYPE DFC_rbr_isobusRegRxDataboxOverlap :
STRUCT
	DTC: UDINT := 16#051100;
	DFCid: UINT := 624;
	debounceMethod: USINT := NO_DEBOUNCE;
END_STRUCT
END_TYPE

(* ---- dfc_rbr_isobusregrxdataboxparam-DFC_rbr_isobusRegRxDataboxParam.st ---- *)
(* --- Interface --- *)
{attribute 'external_name' := 'cmp_rts_DFC_rbr_isobusRegRxDataboxParam'}
TYPE DFC_rbr_isobusRegRxDataboxParam :
STRUCT
	DTC: UDINT := 16#051200;
	DFCid: UINT := 625;
	debounceMethod: USINT := NO_DEBOUNCE;
END_STRUCT
END_TYPE

(* ---- dfc_rbr_isobusregrxdataboxstate-DFC_rbr_isobusRegRxDataboxState.st ---- *)
(* --- Interface --- *)
{attribute 'external_name' := 'cmp_rts_DFC_rbr_isobusRegRxDataboxState'}
TYPE DFC_rbr_isobusRegRxDataboxState :
STRUCT
	DTC: UDINT := 16#051300;
	DFCid: UINT := 626;
	debounceMethod: USINT := NO_DEBOUNCE;
END_STRUCT
END_TYPE

(* ---- dfc_rbr_isobusregtxdataboxoverlap-DFC_rbr_isobusRegTxDataboxOverlap.st ---- *)
(* --- Interface --- *)
{attribute 'external_name' := 'cmp_rts_DFC_rbr_isobusRegTxDataboxOverlap'}
TYPE DFC_rbr_isobusRegTxDataboxOverlap :
STRUCT
	DTC: UDINT := 16#051400;
	DFCid: UINT := 627;
	debounceMethod: USINT := NO_DEBOUNCE;
END_STRUCT
END_TYPE

(* ---- dfc_rbr_isobusregtxdataboxparam-DFC_rbr_isobusRegTxDataboxParam.st ---- *)
(* --- Interface --- *)
{attribute 'external_name' := 'cmp_rts_DFC_rbr_isobusRegTxDataboxParam'}
TYPE DFC_rbr_isobusRegTxDataboxParam :
STRUCT
	DTC: UDINT := 16#051500;
	DFCid: UINT := 628;
	debounceMethod: USINT := NO_DEBOUNCE;
END_STRUCT
END_TYPE

(* ---- dfc_rbr_isobusregtxdataboxstate-DFC_rbr_isobusRegTxDataboxState.st ---- *)
(* --- Interface --- *)
{attribute 'external_name' := 'cmp_rts_DFC_rbr_isobusRegTxDataboxState'}
TYPE DFC_rbr_isobusRegTxDataboxState :
STRUCT
	DTC: UDINT := 16#051600;
	DFCid: UINT := 629;
	debounceMethod: USINT := NO_DEBOUNCE;
END_STRUCT
END_TYPE

(* ---- dfc_rbr_isobussenddataboxparam-DFC_rbr_isobusSendDataboxParam.st ---- *)
(* --- Interface --- *)
{attribute 'external_name' := 'cmp_rts_DFC_rbr_isobusSendDataboxParam'}
TYPE DFC_rbr_isobusSendDataboxParam :
STRUCT
	DTC: UDINT := 16#051700;
	DFCid: UINT := 634;
	debounceMethod: USINT := NO_DEBOUNCE;
END_STRUCT
END_TYPE

(* ---- dfc_rbr_isobussendrequestpgnparam-DFC_rbr_isobusSendRequestPGNParam.st ---- *)
(* --- Interface --- *)
{attribute 'external_name' := 'cmp_rts_DFC_rbr_isobusSendRequestPGNParam'}
TYPE DFC_rbr_isobusSendRequestPGNParam :
STRUCT
	DTC: UDINT := 16#051800;
	DFCid: UINT := 635;
	debounceMethod: USINT := NO_DEBOUNCE;
END_STRUCT
END_TYPE

(* ---- dfc_rbr_isobussetcaaddrcaused-DFC_rbr_isobusSetCaAddrCaUsed.st ---- *)
(* --- Interface --- *)
{attribute 'external_name' := 'cmp_rts_DFC_rbr_isobusSetCaAddrCaUsed'}
TYPE DFC_rbr_isobusSetCaAddrCaUsed :
STRUCT
	DTC: UDINT := 16#051900;
	DFCid: UINT := 636;
	debounceMethod: USINT := NO_DEBOUNCE;
END_STRUCT
END_TYPE

(* ---- dfc_rbr_isobussetcaaddrcomm-DFC_rbr_isobusSetCaAddrComm.st ---- *)
(* --- Interface --- *)
{attribute 'external_name' := 'cmp_rts_DFC_rbr_isobusSetCaAddrComm'}
TYPE DFC_rbr_isobusSetCaAddrComm :
STRUCT
	DTC: UDINT := 16#051A00;
	DFCid: UINT := 637;
	debounceMethod: USINT := NO_DEBOUNCE;
END_STRUCT
END_TYPE

(* ---- dfc_rbr_isobussetcaaddrinvcan-DFC_rbr_isobusSetCaAddrInvCan.st ---- *)
(* --- Interface --- *)
{attribute 'external_name' := 'cmp_rts_DFC_rbr_isobusSetCaAddrInvCan'}
TYPE DFC_rbr_isobusSetCaAddrInvCan :
STRUCT
	DTC: UDINT := 16#051B00;
	DFCid: UINT := 638;
	debounceMethod: USINT := NO_DEBOUNCE;
END_STRUCT
END_TYPE

(* ---- dfc_rbr_isobussetcaaddrparam-DFC_rbr_isobusSetCaAddrParam.st ---- *)
(* --- Interface --- *)
{attribute 'external_name' := 'cmp_rts_DFC_rbr_isobusSetCaAddrParam'}
TYPE DFC_rbr_isobusSetCaAddrParam :
STRUCT
	DTC: UDINT := 16#051C00;
	DFCid: UINT := 639;
	debounceMethod: USINT := NO_DEBOUNCE;
END_STRUCT
END_TYPE

(* ---- dfc_rbr_isobussetcainfoparam-DFC_rbr_isobusSetCaInfoParam.st ---- *)
(* --- Interface --- *)
{attribute 'external_name' := 'cmp_rts_DFC_rbr_isobusSetCaInfoParam'}
TYPE DFC_rbr_isobusSetCaInfoParam :
STRUCT
	DTC: UDINT := 16#051D00;
	DFCid: UINT := 640;
	debounceMethod: USINT := NO_DEBOUNCE;
END_STRUCT
END_TYPE

(* ---- dfc_rbr_isobussetcanameparam-DFC_rbr_isobusSetCaNameParam.st ---- *)
(* --- Interface --- *)
{attribute 'external_name' := 'cmp_rts_DFC_rbr_isobusSetCaNameParam'}
TYPE DFC_rbr_isobusSetCaNameParam :
STRUCT
	DTC: UDINT := 16#051E00;
	DFCid: UINT := 641;
	debounceMethod: USINT := NO_DEBOUNCE;
END_STRUCT
END_TYPE

(* ---- dfc_rbr_isobussftycantxerr-DFC_rbr_isobusSftyCanTxErr.st ---- *)
(* --- Interface --- *)
{attribute 'external_name' := 'cmp_rts_DFC_rbr_isobusSftyCanTxErr'}
TYPE DFC_rbr_isobusSftyCanTxErr :
STRUCT
	DTC: UDINT := 16#051F00;
	DFCid: UINT := 642;
	debounceMethod: USINT := NO_DEBOUNCE;
END_STRUCT
END_TYPE

(* ---- dfc_rbr_lin_getstatus-DFC_rbr_lin_getStatus.st ---- *)
(* --- Interface --- *)
{attribute 'external_name' := 'cmp_rts_DFC_rbr_lin_getStatus'}
TYPE DFC_rbr_lin_getStatus :
STRUCT
	DTC: UDINT := 16#210300;
	DFCid: UINT := 645;
	debounceMethod: USINT := NO_DEBOUNCE;
END_STRUCT
END_TYPE

(* ---- dfc_rbr_lin_gotosleep-DFC_rbr_lin_gotoSleep.st ---- *)
(* --- Interface --- *)
{attribute 'external_name' := 'cmp_rts_DFC_rbr_lin_gotoSleep'}
TYPE DFC_rbr_lin_gotoSleep :
STRUCT
	DTC: UDINT := 16#210200;
	DFCid: UINT := 646;
	debounceMethod: USINT := NO_DEBOUNCE;
END_STRUCT
END_TYPE

(* ---- dfc_rbr_lin_receivesignal-DFC_rbr_lin_ReceiveSignal.st ---- *)
(* --- Interface --- *)
{attribute 'external_name' := 'cmp_rts_DFC_rbr_lin_ReceiveSignal'}
TYPE DFC_rbr_lin_ReceiveSignal :
STRUCT
	DTC: UDINT := 16#210500;
	DFCid: UINT := 643;
	debounceMethod: USINT := NO_DEBOUNCE;
END_STRUCT
END_TYPE

(* ---- dfc_rbr_lin_schedulerequest-DFC_rbr_lin_scheduleRequest.st ---- *)
(* --- Interface --- *)
{attribute 'external_name' := 'cmp_rts_DFC_rbr_lin_scheduleRequest'}
TYPE DFC_rbr_lin_scheduleRequest :
STRUCT
	DTC: UDINT := 16#210100;
	DFCid: UINT := 647;
	debounceMethod: USINT := NO_DEBOUNCE;
END_STRUCT
END_TYPE

(* ---- dfc_rbr_lin_sendsignal-DFC_rbr_lin_SendSignal.st ---- *)
(* --- Interface --- *)
{attribute 'external_name' := 'cmp_rts_DFC_rbr_lin_SendSignal'}
TYPE DFC_rbr_lin_SendSignal :
STRUCT
	DTC: UDINT := 16#210400;
	DFCid: UINT := 644;
	debounceMethod: USINT := NO_DEBOUNCE;
END_STRUCT
END_TYPE

(* ---- dfc_rbr_lin_wakeup-DFC_rbr_lin_wakeUp.st ---- *)
(* --- Interface --- *)
{attribute 'external_name' := 'cmp_rts_DFC_rbr_lin_wakeUp'}
TYPE DFC_rbr_lin_wakeUp :
STRUCT
	DTC: UDINT := 16#210000;
	DFCid: UINT := 648;
	debounceMethod: USINT := NO_DEBOUNCE;
END_STRUCT
END_TYPE

(* ---- dfc_rbr_memflscfgshr-DFC_rbr_memFlsCfgShr.st ---- *)
(* --- Interface --- *)
{attribute 'external_name' := 'cmp_rts_DFC_rbr_memFlsCfgShr'}
TYPE DFC_rbr_memFlsCfgShr :
STRUCT
	DTC: UDINT := 16#060900;
	DFCid: UINT := 649;
	debounceMethod: USINT := NO_DEBOUNCE;
END_STRUCT
END_TYPE

(* ---- dfc_rbr_memgetstatus-DFC_rbr_memGetStatus.st ---- *)
(* --- Interface --- *)
{attribute 'external_name' := 'cmp_rts_DFC_rbr_memGetStatus'}
TYPE DFC_rbr_memGetStatus :
STRUCT
	DTC: UDINT := 16#060300;
	DFCid: UINT := 650;
	debounceMethod: USINT := NO_DEBOUNCE;
END_STRUCT
END_TYPE

(* ---- dfc_rbr_memmarkblock-DFC_rbr_memMarkBlock.st ---- *)
(* --- Interface --- *)
{attribute 'external_name' := 'cmp_rts_DFC_rbr_memMarkBlock'}
TYPE DFC_rbr_memMarkBlock :
STRUCT
	DTC: UDINT := 16#060400;
	DFCid: UINT := 651;
	debounceMethod: USINT := NO_DEBOUNCE;
END_STRUCT
END_TYPE

(* ---- dfc_rbr_memreadapi1error-DFC_rbr_memReadApi1Error.st ---- *)
(* --- Interface --- *)
{attribute 'external_name' := 'cmp_rts_DFC_rbr_memReadApi1Error'}
TYPE DFC_rbr_memReadApi1Error :
STRUCT
	DTC: UDINT := 16#060500;
	DFCid: UINT := 652;
	debounceMethod: USINT := NO_DEBOUNCE;
END_STRUCT
END_TYPE

(* ---- dfc_rbr_memreadapi2error-DFC_rbr_memReadApi2Error.st ---- *)
(* --- Interface --- *)
{attribute 'external_name' := 'cmp_rts_DFC_rbr_memReadApi2Error'}
TYPE DFC_rbr_memReadApi2Error :
STRUCT
	DTC: UDINT := 16#060600;
	DFCid: UINT := 653;
	debounceMethod: USINT := NO_DEBOUNCE;
END_STRUCT
END_TYPE

(* ---- dfc_rbr_memreadblock-DFC_rbr_memReadBlock.st ---- *)
(* --- Interface --- *)
{attribute 'external_name' := 'cmp_rts_DFC_rbr_memReadBlock'}
TYPE DFC_rbr_memReadBlock :
STRUCT
	DTC: UDINT := 16#060200;
	DFCid: UINT := 654;
	debounceMethod: USINT := NO_DEBOUNCE;
END_STRUCT
END_TYPE

(* ---- dfc_rbr_memreadcalibinputerror-DFC_rbr_memReadCalibInputError.st ---- *)
(* --- Interface --- *)
{attribute 'external_name' := 'cmp_rts_DFC_rbr_memReadCalibInputError'}
TYPE DFC_rbr_memReadCalibInputError :
STRUCT
	DTC: UDINT := 16#060A00;
	DFCid: UINT := 655;
	debounceMethod: USINT := NO_DEBOUNCE;
END_STRUCT
END_TYPE

(* ---- dfc_rbr_memreadcalibouputerror-DFC_rbr_memReadCalibOuputError.st ---- *)
(* --- Interface --- *)
{attribute 'external_name' := 'cmp_rts_DFC_rbr_memReadCalibOuputError'}
TYPE DFC_rbr_memReadCalibOuputError :
STRUCT
	DTC: UDINT := 16#060B00;
	DFCid: UINT := 656;
	debounceMethod: USINT := NO_DEBOUNCE;
END_STRUCT
END_TYPE

(* ---- dfc_rbr_memreadsystemerror-DFC_rbr_memReadSystemError.st ---- *)
(* --- Interface --- *)
{attribute 'external_name' := 'cmp_rts_DFC_rbr_memReadSystemError'}
TYPE DFC_rbr_memReadSystemError :
STRUCT
	DTC: UDINT := 16#060800;
	DFCid: UINT := 657;
	debounceMethod: USINT := NO_DEBOUNCE;
END_STRUCT
END_TYPE

(* ---- dfc_rbr_memwriteblock-DFC_rbr_memWriteBlock.st ---- *)
(* --- Interface --- *)
{attribute 'external_name' := 'cmp_rts_DFC_rbr_memWriteBlock'}
TYPE DFC_rbr_memWriteBlock :
STRUCT
	DTC: UDINT := 16#060100;
	DFCid: UINT := 658;
	debounceMethod: USINT := NO_DEBOUNCE;
END_STRUCT
END_TYPE

(* ---- dfc_rbr_mo_adcpdd_fail-DFC_rbr_mo_adcPDD_fail.st ---- *)
(* --- Interface --- *)
{attribute 'external_name' := 'cmp_rts_DFC_rbr_mo_adcPDD_fail'}
TYPE DFC_rbr_mo_adcPDD_fail :
STRUCT
	DTC: UDINT := 16#083000;
	DFCid: UINT := 665;
	debounceMethod: USINT := NO_DEBOUNCE;
END_STRUCT
END_TYPE

(* ---- dfc_rbr_mo_dvubat_fws-DFC_rbr_mo_DvUBAT_FWs.st ---- *)
(* --- Interface --- *)
{attribute 'external_name' := 'cmp_rts_DFC_rbr_mo_DvUBAT_FWs'}
TYPE DFC_rbr_mo_DvUBAT_FWs :
STRUCT
	DTC: UDINT := 16#080D00;
	DFCid: UINT := 243;
	debounceMethod: USINT := TIME_UP_DOWN;
END_STRUCT
END_TYPE

(* ---- dfc_rbr_mo_inh-DFC_rbr_mo_INH.st ---- *)
(* --- Interface --- *)
{attribute 'external_name' := 'cmp_rts_DFC_rbr_mo_INH'}
TYPE DFC_rbr_mo_INH :
STRUCT
	DTC: UDINT := 16#082100;
	DFCid: UINT := 663;
	debounceMethod: USINT := NO_DEBOUNCE;
END_STRUCT
END_TYPE

(* ---- dfc_rbr_mo_inhlatch-DFC_rbr_mo_INHLatch.st ---- *)
(* --- Interface --- *)
{attribute 'external_name' := 'cmp_rts_DFC_rbr_mo_INHLatch'}
TYPE DFC_rbr_mo_INHLatch :
STRUCT
	DTC: UDINT := 16#082200;
	DFCid: UINT := 664;
	debounceMethod: USINT := NO_DEBOUNCE;
END_STRUCT
END_TYPE

(* ---- dfc_rbr_mo_memoryprotection_err-DFC_rbr_mo_memoryProtection_err.st ---- *)
(* --- Interface --- *)
{attribute 'external_name' := 'cmp_rts_DFC_rbr_mo_memoryProtection_err'}
TYPE DFC_rbr_mo_memoryProtection_err :
STRUCT
	DTC: UDINT := 16#083300;
	DFCid: UINT := 666;
	debounceMethod: USINT := NO_DEBOUNCE;
END_STRUCT
END_TYPE

(* ---- dfc_rbr_mo_ov_sav_lss_meas_cluster_1_3-DFC_rbr_mo_OV_SAV_LSS_MEAS_CLUSTER_1_3.st ---- *)
(* --- Interface --- *)
{attribute 'external_name' := 'cmp_rts_DFC_rbr_mo_OV_SAV_LSS_MEAS_CLUSTER_1_3'}
TYPE DFC_rbr_mo_OV_SAV_LSS_MEAS_CLUSTER_1_3 :
STRUCT
	DTC: UDINT := 16#082A00;
	DFCid: UINT := 246;
	debounceMethod: USINT := TIME_UP_DOWN;
END_STRUCT
END_TYPE

(* ---- dfc_rbr_mo_ov_sav_lss_meas_cluster_2-DFC_rbr_mo_OV_SAV_LSS_MEAS_CLUSTER_2.st ---- *)
(* --- Interface --- *)
{attribute 'external_name' := 'cmp_rts_DFC_rbr_mo_OV_SAV_LSS_MEAS_CLUSTER_2'}
TYPE DFC_rbr_mo_OV_SAV_LSS_MEAS_CLUSTER_2 :
STRUCT
	DTC: UDINT := 16#082800;
	DFCid: UINT := 247;
	debounceMethod: USINT := TIME_UP_DOWN;
END_STRUCT
END_TYPE

(* ---- dfc_rbr_mo_ov_ubat_mon-DFC_rbr_mo_OV_UBAT_MON.st ---- *)
(* --- Interface --- *)
{attribute 'external_name' := 'cmp_rts_DFC_rbr_mo_OV_UBAT_MON'}
TYPE DFC_rbr_mo_OV_UBAT_MON :
STRUCT
	DTC: UDINT := 16#080900;
	DFCid: UINT := 248;
	debounceMethod: USINT := TIME_UP_DOWN;
END_STRUCT
END_TYPE

(* ---- dfc_rbr_mo_ov_ubrm24_flexin-DFC_rbr_mo_OV_UBRM24_FLEXIN.st ---- *)
(* --- Interface --- *)
{attribute 'external_name' := 'cmp_rts_DFC_rbr_mo_OV_UBRM24_FLEXIN'}
TYPE DFC_rbr_mo_OV_UBRM24_FLEXIN :
STRUCT
	DTC: UDINT := 16#082300;
	DFCid: UINT := 249;
	debounceMethod: USINT := TIME_UP_DOWN;
END_STRUCT
END_TYPE

(* ---- dfc_rbr_mo_ov_ubrm24_loads-DFC_rbr_mo_OV_UBRM24_LOADS.st ---- *)
(* --- Interface --- *)
{attribute 'external_name' := 'cmp_rts_DFC_rbr_mo_OV_UBRM24_LOADS'}
TYPE DFC_rbr_mo_OV_UBRM24_LOADS :
STRUCT
	DTC: UDINT := 16#080C00;
	DFCid: UINT := 250;
	debounceMethod: USINT := TIME_UP_DOWN;
END_STRUCT
END_TYPE

(* ---- dfc_rbr_mo_ov_ubrm24_mon-DFC_rbr_mo_OV_UBRM24_MON.st ---- *)
(* --- Interface --- *)
{attribute 'external_name' := 'cmp_rts_DFC_rbr_mo_OV_UBRM24_MON'}
TYPE DFC_rbr_mo_OV_UBRM24_MON :
STRUCT
	DTC: UDINT := 16#080A00;
	DFCid: UINT := 251;
	debounceMethod: USINT := TIME_UP_DOWN;
END_STRUCT
END_TYPE

(* ---- dfc_rbr_mo_ov_vdd5-DFC_rbr_mo_OV_VDD5.st ---- *)
(* --- Interface --- *)
{attribute 'external_name' := 'cmp_rts_DFC_rbr_mo_OV_VDD5'}
TYPE DFC_rbr_mo_OV_VDD5 :
STRUCT
	DTC: UDINT := 16#082400;
	DFCid: UINT := 252;
	debounceMethod: USINT := TIME_UP_DOWN;
END_STRUCT
END_TYPE

(* ---- dfc_rbr_mo_ov_vdd5_in-DFC_rbr_mo_OV_VDD5_IN.st ---- *)
(* --- Interface --- *)
{attribute 'external_name' := 'cmp_rts_DFC_rbr_mo_OV_VDD5_IN'}
TYPE DFC_rbr_mo_OV_VDD5_IN :
STRUCT
	DTC: UDINT := 16#082600;
	DFCid: UINT := 253;
	debounceMethod: USINT := TIME_UP_DOWN;
END_STRUCT
END_TYPE

(* ---- dfc_rbr_mo_ov_vpr6-DFC_rbr_mo_OV_VPR6.st ---- *)
(* --- Interface --- *)
{attribute 'external_name' := 'cmp_rts_DFC_rbr_mo_OV_VPR6'}
TYPE DFC_rbr_mo_OV_VPR6 :
STRUCT
	DTC: UDINT := 16#082000;
	DFCid: UINT := 254;
	debounceMethod: USINT := TIME_UP_DOWN;
END_STRUCT
END_TYPE

(* ---- dfc_rbr_mo_ov_vss1-DFC_rbr_mo_OV_VSS1.st ---- *)
(* --- Interface --- *)
{attribute 'external_name' := 'cmp_rts_DFC_rbr_mo_OV_VSS1'}
TYPE DFC_rbr_mo_OV_VSS1 :
STRUCT
	DTC: UDINT := 16#080100;
	DFCid: UINT := 852;
	debounceMethod: USINT := NO_DEBOUNCE;
END_STRUCT
END_TYPE

(* ---- dfc_rbr_mo_ov_vss2-DFC_rbr_mo_OV_VSS2.st ---- *)
(* --- Interface --- *)
{attribute 'external_name' := 'cmp_rts_DFC_rbr_mo_OV_VSS2'}
TYPE DFC_rbr_mo_OV_VSS2 :
STRUCT
	DTC: UDINT := 16#080300;
	DFCid: UINT := 853;
	debounceMethod: USINT := NO_DEBOUNCE;
END_STRUCT
END_TYPE

(* ---- dfc_rbr_mo_ov_vss3-DFC_rbr_mo_OV_VSS3.st ---- *)
(* --- Interface --- *)
{attribute 'external_name' := 'cmp_rts_DFC_rbr_mo_OV_VSS3'}
TYPE DFC_rbr_mo_OV_VSS3 :
STRUCT
	DTC: UDINT := 16#080500;
	DFCid: UINT := 255;
	debounceMethod: USINT := TIME_UP_DOWN;
END_STRUCT
END_TYPE

(* ---- dfc_rbr_mo_ov_vss4-DFC_rbr_mo_OV_VSS4.st ---- *)
(* --- Interface --- *)
{attribute 'external_name' := 'cmp_rts_DFC_rbr_mo_OV_VSS4'}
TYPE DFC_rbr_mo_OV_VSS4 :
STRUCT
	DTC: UDINT := 16#080700;
	DFCid: UINT := 256;
	debounceMethod: USINT := TIME_UP_DOWN;
END_STRUCT
END_TYPE

(* ---- dfc_rbr_mo_overr_vpr6-DFC_rbr_mo_OVErr_VPR6.st ---- *)
(* --- Interface --- *)
{attribute 'external_name' := 'cmp_rts_DFC_rbr_mo_OVErr_VPR6'}
TYPE DFC_rbr_mo_OVErr_VPR6 :
STRUCT
	DTC: UDINT := 16#081100;
	DFCid: UINT := 244;
	debounceMethod: USINT := TIME_UP_DOWN;
END_STRUCT
END_TYPE

(* ---- dfc_rbr_mo_ovwarn_vpr6-DFC_rbr_mo_OVWarn_VPR6.st ---- *)
(* --- Interface --- *)
{attribute 'external_name' := 'cmp_rts_DFC_rbr_mo_OVWarn_VPR6'}
TYPE DFC_rbr_mo_OVWarn_VPR6 :
STRUCT
	DTC: UDINT := 16#081200;
	DFCid: UINT := 245;
	debounceMethod: USINT := TIME_UP_DOWN;
END_STRUCT
END_TYPE

(* ---- dfc_rbr_mo_temp1_hterr-DFC_rbr_mo_Temp1_HTErr.st ---- *)
(* --- Interface --- *)
{attribute 'external_name' := 'cmp_rts_DFC_rbr_mo_Temp1_HTErr'}
TYPE DFC_rbr_mo_Temp1_HTErr :
STRUCT
	DTC: UDINT := 16#081700;
	DFCid: UINT := 257;
	debounceMethod: USINT := TIME_UP_DOWN;
END_STRUCT
END_TYPE

(* ---- dfc_rbr_mo_temp1_htwarn-DFC_rbr_mo_Temp1_HTWarn.st ---- *)
(* --- Interface --- *)
{attribute 'external_name' := 'cmp_rts_DFC_rbr_mo_Temp1_HTWarn'}
TYPE DFC_rbr_mo_Temp1_HTWarn :
STRUCT
	DTC: UDINT := 16#081600;
	DFCid: UINT := 258;
	debounceMethod: USINT := TIME_UP_DOWN;
END_STRUCT
END_TYPE

(* ---- dfc_rbr_mo_temp2_hterr-DFC_rbr_mo_Temp2_HTErr.st ---- *)
(* --- Interface --- *)
{attribute 'external_name' := 'cmp_rts_DFC_rbr_mo_Temp2_HTErr'}
TYPE DFC_rbr_mo_Temp2_HTErr :
STRUCT
	DTC: UDINT := 16#081900;
	DFCid: UINT := 259;
	debounceMethod: USINT := TIME_UP_DOWN;
END_STRUCT
END_TYPE

(* ---- dfc_rbr_mo_temp2_htwarn-DFC_rbr_mo_Temp2_HTWarn.st ---- *)
(* --- Interface --- *)
{attribute 'external_name' := 'cmp_rts_DFC_rbr_mo_Temp2_HTWarn'}
TYPE DFC_rbr_mo_Temp2_HTWarn :
STRUCT
	DTC: UDINT := 16#081800;
	DFCid: UINT := 260;
	debounceMethod: USINT := TIME_UP_DOWN;
END_STRUCT
END_TYPE

(* ---- dfc_rbr_mo_uv_sav_lss_meas_cluster_1_3-DFC_rbr_mo_UV_SAV_LSS_MEAS_CLUSTER_1_3.st ---- *)
(* --- Interface --- *)
{attribute 'external_name' := 'cmp_rts_DFC_rbr_mo_UV_SAV_LSS_MEAS_CLUSTER_1_3'}
TYPE DFC_rbr_mo_UV_SAV_LSS_MEAS_CLUSTER_1_3 :
STRUCT
	DTC: UDINT := 16#082B00;
	DFCid: UINT := 261;
	debounceMethod: USINT := TIME_UP_DOWN;
END_STRUCT
END_TYPE

(* ---- dfc_rbr_mo_uv_sav_lss_meas_cluster_2-DFC_rbr_mo_UV_SAV_LSS_MEAS_CLUSTER_2.st ---- *)
(* --- Interface --- *)
{attribute 'external_name' := 'cmp_rts_DFC_rbr_mo_UV_SAV_LSS_MEAS_CLUSTER_2'}
TYPE DFC_rbr_mo_UV_SAV_LSS_MEAS_CLUSTER_2 :
STRUCT
	DTC: UDINT := 16#082900;
	DFCid: UINT := 262;
	debounceMethod: USINT := TIME_UP_DOWN;
END_STRUCT
END_TYPE

(* ---- dfc_rbr_mo_uv_vdd5-DFC_rbr_mo_UV_VDD5.st ---- *)
(* --- Interface --- *)
{attribute 'external_name' := 'cmp_rts_DFC_rbr_mo_UV_VDD5'}
TYPE DFC_rbr_mo_UV_VDD5 :
STRUCT
	DTC: UDINT := 16#082500;
	DFCid: UINT := 263;
	debounceMethod: USINT := TIME_UP_DOWN;
END_STRUCT
END_TYPE

(* ---- dfc_rbr_mo_uv_vdd5_in-DFC_rbr_mo_UV_VDD5_IN.st ---- *)
(* --- Interface --- *)
{attribute 'external_name' := 'cmp_rts_DFC_rbr_mo_UV_VDD5_IN'}
TYPE DFC_rbr_mo_UV_VDD5_IN :
STRUCT
	DTC: UDINT := 16#082700;
	DFCid: UINT := 264;
	debounceMethod: USINT := TIME_UP_DOWN;
END_STRUCT
END_TYPE

(* ---- dfc_rbr_mo_uv_vpr6-DFC_rbr_mo_UV_VPR6.st ---- *)
(* --- Interface --- *)
{attribute 'external_name' := 'cmp_rts_DFC_rbr_mo_UV_VPR6'}
TYPE DFC_rbr_mo_UV_VPR6 :
STRUCT
	DTC: UDINT := 16#081300;
	DFCid: UINT := 265;
	debounceMethod: USINT := TIME_UP_DOWN;
END_STRUCT
END_TYPE

(* ---- dfc_rbr_mo_uv_vss1-DFC_rbr_mo_UV_VSS1.st ---- *)
(* --- Interface --- *)
{attribute 'external_name' := 'cmp_rts_DFC_rbr_mo_UV_VSS1'}
TYPE DFC_rbr_mo_UV_VSS1 :
STRUCT
	DTC: UDINT := 16#080200;
	DFCid: UINT := 854;
	debounceMethod: USINT := NO_DEBOUNCE;
END_STRUCT
END_TYPE

(* ---- dfc_rbr_mo_uv_vss2-DFC_rbr_mo_UV_VSS2.st ---- *)
(* --- Interface --- *)
{attribute 'external_name' := 'cmp_rts_DFC_rbr_mo_UV_VSS2'}
TYPE DFC_rbr_mo_UV_VSS2 :
STRUCT
	DTC: UDINT := 16#080400;
	DFCid: UINT := 855;
	debounceMethod: USINT := NO_DEBOUNCE;
END_STRUCT
END_TYPE

(* ---- dfc_rbr_mo_uv_vss3-DFC_rbr_mo_UV_VSS3.st ---- *)
(* --- Interface --- *)
{attribute 'external_name' := 'cmp_rts_DFC_rbr_mo_UV_VSS3'}
TYPE DFC_rbr_mo_UV_VSS3 :
STRUCT
	DTC: UDINT := 16#080600;
	DFCid: UINT := 266;
	debounceMethod: USINT := TIME_UP_DOWN;
END_STRUCT
END_TYPE

(* ---- dfc_rbr_mo_uv_vss4-DFC_rbr_mo_UV_VSS4.st ---- *)
(* --- Interface --- *)
{attribute 'external_name' := 'cmp_rts_DFC_rbr_mo_UV_VSS4'}
TYPE DFC_rbr_mo_UV_VSS4 :
STRUCT
	DTC: UDINT := 16#080800;
	DFCid: UINT := 267;
	debounceMethod: USINT := TIME_UP_DOWN;
END_STRUCT
END_TYPE

(* ---- dfc_rbr_moov_firstconstadc-DFC_rbr_moOV_FirstConstADC.st ---- *)
(* --- Interface --- *)
{attribute 'external_name' := 'cmp_rts_DFC_rbr_moOV_FirstConstADC'}
TYPE DFC_rbr_moOV_FirstConstADC :
STRUCT
	DTC: UDINT := 16#082C00;
	DFCid: UINT := 659;
	debounceMethod: USINT := NO_DEBOUNCE;
END_STRUCT
END_TYPE

(* ---- dfc_rbr_moov_secondconstadc-DFC_rbr_moOV_SecondConstADC.st ---- *)
(* --- Interface --- *)
{attribute 'external_name' := 'cmp_rts_DFC_rbr_moOV_SecondConstADC'}
TYPE DFC_rbr_moOV_SecondConstADC :
STRUCT
	DTC: UDINT := 16#082E00;
	DFCid: UINT := 660;
	debounceMethod: USINT := NO_DEBOUNCE;
END_STRUCT
END_TYPE

(* ---- dfc_rbr_mouv_firstconstadc-DFC_rbr_moUV_FirstConstADC.st ---- *)
(* --- Interface --- *)
{attribute 'external_name' := 'cmp_rts_DFC_rbr_moUV_FirstConstADC'}
TYPE DFC_rbr_moUV_FirstConstADC :
STRUCT
	DTC: UDINT := 16#082D00;
	DFCid: UINT := 661;
	debounceMethod: USINT := NO_DEBOUNCE;
END_STRUCT
END_TYPE

(* ---- dfc_rbr_mouv_secondconstadc-DFC_rbr_moUV_SecondConstADC.st ---- *)
(* --- Interface --- *)
{attribute 'external_name' := 'cmp_rts_DFC_rbr_moUV_SecondConstADC'}
TYPE DFC_rbr_moUV_SecondConstADC :
STRUCT
	DTC: UDINT := 16#082F00;
	DFCid: UINT := 662;
	debounceMethod: USINT := NO_DEBOUNCE;
END_STRUCT
END_TYPE

(* ---- dfc_rbr_outa01ol-DFC_rbr_outA01OL.st ---- *)
(* --- Interface --- *)
{attribute 'external_name' := 'cmp_rts_DFC_rbr_outA01OL'}
TYPE DFC_rbr_outA01OL :
STRUCT
	DTC: UDINT := 16#140100;
	DFCid: UINT := 268;
	debounceMethod: USINT := TIME_UP_DOWN;
END_STRUCT
END_TYPE

(* ---- dfc_rbr_outa01ot-DFC_rbr_outA01OT.st ---- *)
(* --- Interface --- *)
{attribute 'external_name' := 'cmp_rts_DFC_rbr_outA01OT'}
TYPE DFC_rbr_outA01OT :
STRUCT
	DTC: UDINT := 16#140200;
	DFCid: UINT := 269;
	debounceMethod: USINT := TIME_UP_DOWN;
END_STRUCT
END_TYPE

(* ---- dfc_rbr_outa01scb-DFC_rbr_outA01SCB.st ---- *)
(* --- Interface --- *)
{attribute 'external_name' := 'cmp_rts_DFC_rbr_outA01SCB'}
TYPE DFC_rbr_outA01SCB :
STRUCT
	DTC: UDINT := 16#140300;
	DFCid: UINT := 270;
	debounceMethod: USINT := TIME_UP_DOWN;
END_STRUCT
END_TYPE

(* ---- dfc_rbr_outa01scg-DFC_rbr_outA01SCG.st ---- *)
(* --- Interface --- *)
{attribute 'external_name' := 'cmp_rts_DFC_rbr_outA01SCG'}
TYPE DFC_rbr_outA01SCG :
STRUCT
	DTC: UDINT := 16#140400;
	DFCid: UINT := 271;
	debounceMethod: USINT := TIME_UP_DOWN;
END_STRUCT
END_TYPE

(* ---- dfc_rbr_outa02oc-DFC_rbr_outA02OC.st ---- *)
(* --- Interface --- *)
{attribute 'external_name' := 'cmp_rts_DFC_rbr_outA02OC'}
TYPE DFC_rbr_outA02OC :
STRUCT
	DTC: UDINT := 16#140500;
	DFCid: UINT := 667;
	debounceMethod: USINT := NO_DEBOUNCE;
END_STRUCT
END_TYPE

(* ---- dfc_rbr_outa02ol-DFC_rbr_outA02OL.st ---- *)
(* --- Interface --- *)
{attribute 'external_name' := 'cmp_rts_DFC_rbr_outA02OL'}
TYPE DFC_rbr_outA02OL :
STRUCT
	DTC: UDINT := 16#140600;
	DFCid: UINT := 272;
	debounceMethod: USINT := TIME_UP_DOWN;
END_STRUCT
END_TYPE

(* ---- dfc_rbr_outa02or-DFC_rbr_outA02OR.st ---- *)
(* --- Interface --- *)
{attribute 'external_name' := 'cmp_rts_DFC_rbr_outA02OR'}
TYPE DFC_rbr_outA02OR :
STRUCT
	DTC: UDINT := 16#140700;
	DFCid: UINT := 273;
	debounceMethod: USINT := TIME_UP_DOWN;
END_STRUCT
END_TYPE

(* ---- dfc_rbr_outa02ot-DFC_rbr_outA02OT.st ---- *)
(* --- Interface --- *)
{attribute 'external_name' := 'cmp_rts_DFC_rbr_outA02OT'}
TYPE DFC_rbr_outA02OT :
STRUCT
	DTC: UDINT := 16#140800;
	DFCid: UINT := 274;
	debounceMethod: USINT := TIME_UP_DOWN;
END_STRUCT
END_TYPE

(* ---- dfc_rbr_outa02scb-DFC_rbr_outA02SCB.st ---- *)
(* --- Interface --- *)
{attribute 'external_name' := 'cmp_rts_DFC_rbr_outA02SCB'}
TYPE DFC_rbr_outA02SCB :
STRUCT
	DTC: UDINT := 16#140900;
	DFCid: UINT := 275;
	debounceMethod: USINT := TIME_UP_DOWN;
END_STRUCT
END_TYPE

(* ---- dfc_rbr_outa02scg-DFC_rbr_outA02SCG.st ---- *)
(* --- Interface --- *)
{attribute 'external_name' := 'cmp_rts_DFC_rbr_outA02SCG'}
TYPE DFC_rbr_outA02SCG :
STRUCT
	DTC: UDINT := 16#140A00;
	DFCid: UINT := 276;
	debounceMethod: USINT := TIME_UP_DOWN;
END_STRUCT
END_TYPE

(* ---- dfc_rbr_outa02unintended-DFC_rbr_outA02Unintended.st ---- *)
(* --- Interface --- *)
{attribute 'external_name' := 'cmp_rts_DFC_rbr_outA02Unintended'}
TYPE DFC_rbr_outA02Unintended :
STRUCT
	DTC: UDINT := 16#14B300;
	DFCid: UINT := 668;
	debounceMethod: USINT := NO_DEBOUNCE;
END_STRUCT
END_TYPE

(* ---- dfc_rbr_outa03oc-DFC_rbr_outA03OC.st ---- *)
(* --- Interface --- *)
{attribute 'external_name' := 'cmp_rts_DFC_rbr_outA03OC'}
TYPE DFC_rbr_outA03OC :
STRUCT
	DTC: UDINT := 16#140B00;
	DFCid: UINT := 669;
	debounceMethod: USINT := NO_DEBOUNCE;
END_STRUCT
END_TYPE

(* ---- dfc_rbr_outa03ol-DFC_rbr_outA03OL.st ---- *)
(* --- Interface --- *)
{attribute 'external_name' := 'cmp_rts_DFC_rbr_outA03OL'}
TYPE DFC_rbr_outA03OL :
STRUCT
	DTC: UDINT := 16#140C00;
	DFCid: UINT := 277;
	debounceMethod: USINT := TIME_UP_DOWN;
END_STRUCT
END_TYPE

(* ---- dfc_rbr_outa03ot-DFC_rbr_outA03OT.st ---- *)
(* --- Interface --- *)
{attribute 'external_name' := 'cmp_rts_DFC_rbr_outA03OT'}
TYPE DFC_rbr_outA03OT :
STRUCT
	DTC: UDINT := 16#140D00;
	DFCid: UINT := 278;
	debounceMethod: USINT := TIME_UP_DOWN;
END_STRUCT
END_TYPE

(* ---- dfc_rbr_outa03scb-DFC_rbr_outA03SCB.st ---- *)
(* --- Interface --- *)
{attribute 'external_name' := 'cmp_rts_DFC_rbr_outA03SCB'}
TYPE DFC_rbr_outA03SCB :
STRUCT
	DTC: UDINT := 16#140E00;
	DFCid: UINT := 279;
	debounceMethod: USINT := TIME_UP_DOWN;
END_STRUCT
END_TYPE

(* ---- dfc_rbr_outa03scg-DFC_rbr_outA03SCG.st ---- *)
(* --- Interface --- *)
{attribute 'external_name' := 'cmp_rts_DFC_rbr_outA03SCG'}
TYPE DFC_rbr_outA03SCG :
STRUCT
	DTC: UDINT := 16#140F00;
	DFCid: UINT := 280;
	debounceMethod: USINT := TIME_UP_DOWN;
END_STRUCT
END_TYPE

(* ---- dfc_rbr_outa03unintended-DFC_rbr_outA03Unintended.st ---- *)
(* --- Interface --- *)
{attribute 'external_name' := 'cmp_rts_DFC_rbr_outA03Unintended'}
TYPE DFC_rbr_outA03Unintended :
STRUCT
	DTC: UDINT := 16#14B400;
	DFCid: UINT := 670;
	debounceMethod: USINT := NO_DEBOUNCE;
END_STRUCT
END_TYPE

(* ---- dfc_rbr_outa04oc-DFC_rbr_outA04OC.st ---- *)
(* --- Interface --- *)
{attribute 'external_name' := 'cmp_rts_DFC_rbr_outA04OC'}
TYPE DFC_rbr_outA04OC :
STRUCT
	DTC: UDINT := 16#141000;
	DFCid: UINT := 671;
	debounceMethod: USINT := NO_DEBOUNCE;
END_STRUCT
END_TYPE

(* ---- dfc_rbr_outa04ol-DFC_rbr_outA04OL.st ---- *)
(* --- Interface --- *)
{attribute 'external_name' := 'cmp_rts_DFC_rbr_outA04OL'}
TYPE DFC_rbr_outA04OL :
STRUCT
	DTC: UDINT := 16#141100;
	DFCid: UINT := 281;
	debounceMethod: USINT := TIME_UP_DOWN;
END_STRUCT
END_TYPE

(* ---- dfc_rbr_outa04ot-DFC_rbr_outA04OT.st ---- *)
(* --- Interface --- *)
{attribute 'external_name' := 'cmp_rts_DFC_rbr_outA04OT'}
TYPE DFC_rbr_outA04OT :
STRUCT
	DTC: UDINT := 16#141200;
	DFCid: UINT := 282;
	debounceMethod: USINT := TIME_UP_DOWN;
END_STRUCT
END_TYPE

(* ---- dfc_rbr_outa04scb-DFC_rbr_outA04SCB.st ---- *)
(* --- Interface --- *)
{attribute 'external_name' := 'cmp_rts_DFC_rbr_outA04SCB'}
TYPE DFC_rbr_outA04SCB :
STRUCT
	DTC: UDINT := 16#141300;
	DFCid: UINT := 283;
	debounceMethod: USINT := TIME_UP_DOWN;
END_STRUCT
END_TYPE

(* ---- dfc_rbr_outa04scg-DFC_rbr_outA04SCG.st ---- *)
(* --- Interface --- *)
{attribute 'external_name' := 'cmp_rts_DFC_rbr_outA04SCG'}
TYPE DFC_rbr_outA04SCG :
STRUCT
	DTC: UDINT := 16#141400;
	DFCid: UINT := 284;
	debounceMethod: USINT := TIME_UP_DOWN;
END_STRUCT
END_TYPE

(* ---- dfc_rbr_outa04unintended-DFC_rbr_outA04Unintended.st ---- *)
(* --- Interface --- *)
{attribute 'external_name' := 'cmp_rts_DFC_rbr_outA04Unintended'}
TYPE DFC_rbr_outA04Unintended :
STRUCT
	DTC: UDINT := 16#14B500;
	DFCid: UINT := 672;
	debounceMethod: USINT := NO_DEBOUNCE;
END_STRUCT
END_TYPE

(* ---- dfc_rbr_outa05oc-DFC_rbr_outA05OC.st ---- *)
(* --- Interface --- *)
{attribute 'external_name' := 'cmp_rts_DFC_rbr_outA05OC'}
TYPE DFC_rbr_outA05OC :
STRUCT
	DTC: UDINT := 16#141500;
	DFCid: UINT := 673;
	debounceMethod: USINT := NO_DEBOUNCE;
END_STRUCT
END_TYPE

(* ---- dfc_rbr_outa05ol-DFC_rbr_outA05OL.st ---- *)
(* --- Interface --- *)
{attribute 'external_name' := 'cmp_rts_DFC_rbr_outA05OL'}
TYPE DFC_rbr_outA05OL :
STRUCT
	DTC: UDINT := 16#141600;
	DFCid: UINT := 285;
	debounceMethod: USINT := TIME_UP_DOWN;
END_STRUCT
END_TYPE

(* ---- dfc_rbr_outa05or-DFC_rbr_outA05OR.st ---- *)
(* --- Interface --- *)
{attribute 'external_name' := 'cmp_rts_DFC_rbr_outA05OR'}
TYPE DFC_rbr_outA05OR :
STRUCT
	DTC: UDINT := 16#141700;
	DFCid: UINT := 286;
	debounceMethod: USINT := TIME_UP_DOWN;
END_STRUCT
END_TYPE

(* ---- dfc_rbr_outa05ot-DFC_rbr_outA05OT.st ---- *)
(* --- Interface --- *)
{attribute 'external_name' := 'cmp_rts_DFC_rbr_outA05OT'}
TYPE DFC_rbr_outA05OT :
STRUCT
	DTC: UDINT := 16#141800;
	DFCid: UINT := 287;
	debounceMethod: USINT := TIME_UP_DOWN;
END_STRUCT
END_TYPE

(* ---- dfc_rbr_outa05scb-DFC_rbr_outA05SCB.st ---- *)
(* --- Interface --- *)
{attribute 'external_name' := 'cmp_rts_DFC_rbr_outA05SCB'}
TYPE DFC_rbr_outA05SCB :
STRUCT
	DTC: UDINT := 16#141900;
	DFCid: UINT := 288;
	debounceMethod: USINT := TIME_UP_DOWN;
END_STRUCT
END_TYPE

(* ---- dfc_rbr_outa05scg-DFC_rbr_outA05SCG.st ---- *)
(* --- Interface --- *)
{attribute 'external_name' := 'cmp_rts_DFC_rbr_outA05SCG'}
TYPE DFC_rbr_outA05SCG :
STRUCT
	DTC: UDINT := 16#141A00;
	DFCid: UINT := 289;
	debounceMethod: USINT := TIME_UP_DOWN;
END_STRUCT
END_TYPE

(* ---- dfc_rbr_outa05unintended-DFC_rbr_outA05Unintended.st ---- *)
(* --- Interface --- *)
{attribute 'external_name' := 'cmp_rts_DFC_rbr_outA05Unintended'}
TYPE DFC_rbr_outA05Unintended :
STRUCT
	DTC: UDINT := 16#14B600;
	DFCid: UINT := 674;
	debounceMethod: USINT := NO_DEBOUNCE;
END_STRUCT
END_TYPE

(* ---- dfc_rbr_outa06ol-DFC_rbr_outA06OL.st ---- *)
(* --- Interface --- *)
{attribute 'external_name' := 'cmp_rts_DFC_rbr_outA06OL'}
TYPE DFC_rbr_outA06OL :
STRUCT
	DTC: UDINT := 16#141B00;
	DFCid: UINT := 290;
	debounceMethod: USINT := TIME_UP_DOWN;
END_STRUCT
END_TYPE

(* ---- dfc_rbr_outa06or-DFC_rbr_outA06OR.st ---- *)
(* --- Interface --- *)
{attribute 'external_name' := 'cmp_rts_DFC_rbr_outA06OR'}
TYPE DFC_rbr_outA06OR :
STRUCT
	DTC: UDINT := 16#141C00;
	DFCid: UINT := 291;
	debounceMethod: USINT := TIME_UP_DOWN;
END_STRUCT
END_TYPE

(* ---- dfc_rbr_outa06ot-DFC_rbr_outA06OT.st ---- *)
(* --- Interface --- *)
{attribute 'external_name' := 'cmp_rts_DFC_rbr_outA06OT'}
TYPE DFC_rbr_outA06OT :
STRUCT
	DTC: UDINT := 16#141D00;
	DFCid: UINT := 292;
	debounceMethod: USINT := TIME_UP_DOWN;
END_STRUCT
END_TYPE

(* ---- dfc_rbr_outa06scb-DFC_rbr_outA06SCB.st ---- *)
(* --- Interface --- *)
{attribute 'external_name' := 'cmp_rts_DFC_rbr_outA06SCB'}
TYPE DFC_rbr_outA06SCB :
STRUCT
	DTC: UDINT := 16#141E00;
	DFCid: UINT := 293;
	debounceMethod: USINT := TIME_UP_DOWN;
END_STRUCT
END_TYPE

(* ---- dfc_rbr_outa06scg-DFC_rbr_outA06SCG.st ---- *)
(* --- Interface --- *)
{attribute 'external_name' := 'cmp_rts_DFC_rbr_outA06SCG'}
TYPE DFC_rbr_outA06SCG :
STRUCT
	DTC: UDINT := 16#141F00;
	DFCid: UINT := 294;
	debounceMethod: USINT := TIME_UP_DOWN;
END_STRUCT
END_TYPE

(* ---- dfc_rbr_outa07oc-DFC_rbr_outA07OC.st ---- *)
(* --- Interface --- *)
{attribute 'external_name' := 'cmp_rts_DFC_rbr_outA07OC'}
TYPE DFC_rbr_outA07OC :
STRUCT
	DTC: UDINT := 16#142000;
	DFCid: UINT := 675;
	debounceMethod: USINT := NO_DEBOUNCE;
END_STRUCT
END_TYPE

(* ---- dfc_rbr_outa07ol-DFC_rbr_outA07OL.st ---- *)
(* --- Interface --- *)
{attribute 'external_name' := 'cmp_rts_DFC_rbr_outA07OL'}
TYPE DFC_rbr_outA07OL :
STRUCT
	DTC: UDINT := 16#142100;
	DFCid: UINT := 295;
	debounceMethod: USINT := TIME_UP_DOWN;
END_STRUCT
END_TYPE

(* ---- dfc_rbr_outa07ot-DFC_rbr_outA07OT.st ---- *)
(* --- Interface --- *)
{attribute 'external_name' := 'cmp_rts_DFC_rbr_outA07OT'}
TYPE DFC_rbr_outA07OT :
STRUCT
	DTC: UDINT := 16#142200;
	DFCid: UINT := 296;
	debounceMethod: USINT := TIME_UP_DOWN;
END_STRUCT
END_TYPE

(* ---- dfc_rbr_outa07scb-DFC_rbr_outA07SCB.st ---- *)
(* --- Interface --- *)
{attribute 'external_name' := 'cmp_rts_DFC_rbr_outA07SCB'}
TYPE DFC_rbr_outA07SCB :
STRUCT
	DTC: UDINT := 16#142300;
	DFCid: UINT := 297;
	debounceMethod: USINT := TIME_UP_DOWN;
END_STRUCT
END_TYPE

(* ---- dfc_rbr_outa07scg-DFC_rbr_outA07SCG.st ---- *)
(* --- Interface --- *)
{attribute 'external_name' := 'cmp_rts_DFC_rbr_outA07SCG'}
TYPE DFC_rbr_outA07SCG :
STRUCT
	DTC: UDINT := 16#142400;
	DFCid: UINT := 298;
	debounceMethod: USINT := TIME_UP_DOWN;
END_STRUCT
END_TYPE

(* ---- dfc_rbr_outa07unintended-DFC_rbr_outA07Unintended.st ---- *)
(* --- Interface --- *)
{attribute 'external_name' := 'cmp_rts_DFC_rbr_outA07Unintended'}
TYPE DFC_rbr_outA07Unintended :
STRUCT
	DTC: UDINT := 16#14B700;
	DFCid: UINT := 676;
	debounceMethod: USINT := NO_DEBOUNCE;
END_STRUCT
END_TYPE

(* ---- dfc_rbr_outa08oc-DFC_rbr_outA08OC.st ---- *)
(* --- Interface --- *)
{attribute 'external_name' := 'cmp_rts_DFC_rbr_outA08OC'}
TYPE DFC_rbr_outA08OC :
STRUCT
	DTC: UDINT := 16#142500;
	DFCid: UINT := 677;
	debounceMethod: USINT := NO_DEBOUNCE;
END_STRUCT
END_TYPE

(* ---- dfc_rbr_outa08ol-DFC_rbr_outA08OL.st ---- *)
(* --- Interface --- *)
{attribute 'external_name' := 'cmp_rts_DFC_rbr_outA08OL'}
TYPE DFC_rbr_outA08OL :
STRUCT
	DTC: UDINT := 16#142600;
	DFCid: UINT := 299;
	debounceMethod: USINT := TIME_UP_DOWN;
END_STRUCT
END_TYPE

(* ---- dfc_rbr_outa08ot-DFC_rbr_outA08OT.st ---- *)
(* --- Interface --- *)
{attribute 'external_name' := 'cmp_rts_DFC_rbr_outA08OT'}
TYPE DFC_rbr_outA08OT :
STRUCT
	DTC: UDINT := 16#142700;
	DFCid: UINT := 300;
	debounceMethod: USINT := TIME_UP_DOWN;
END_STRUCT
END_TYPE

(* ---- dfc_rbr_outa08scb-DFC_rbr_outA08SCB.st ---- *)
(* --- Interface --- *)
{attribute 'external_name' := 'cmp_rts_DFC_rbr_outA08SCB'}
TYPE DFC_rbr_outA08SCB :
STRUCT
	DTC: UDINT := 16#142800;
	DFCid: UINT := 301;
	debounceMethod: USINT := TIME_UP_DOWN;
END_STRUCT
END_TYPE

(* ---- dfc_rbr_outa08scg-DFC_rbr_outA08SCG.st ---- *)
(* --- Interface --- *)
{attribute 'external_name' := 'cmp_rts_DFC_rbr_outA08SCG'}
TYPE DFC_rbr_outA08SCG :
STRUCT
	DTC: UDINT := 16#142900;
	DFCid: UINT := 302;
	debounceMethod: USINT := TIME_UP_DOWN;
END_STRUCT
END_TYPE

(* ---- dfc_rbr_outa08unintended-DFC_rbr_outA08Unintended.st ---- *)
(* --- Interface --- *)
{attribute 'external_name' := 'cmp_rts_DFC_rbr_outA08Unintended'}
TYPE DFC_rbr_outA08Unintended :
STRUCT
	DTC: UDINT := 16#14B800;
	DFCid: UINT := 678;
	debounceMethod: USINT := NO_DEBOUNCE;
END_STRUCT
END_TYPE

(* ---- dfc_rbr_outa09oc-DFC_rbr_outA09OC.st ---- *)
(* --- Interface --- *)
{attribute 'external_name' := 'cmp_rts_DFC_rbr_outA09OC'}
TYPE DFC_rbr_outA09OC :
STRUCT
	DTC: UDINT := 16#142A00;
	DFCid: UINT := 679;
	debounceMethod: USINT := NO_DEBOUNCE;
END_STRUCT
END_TYPE

(* ---- dfc_rbr_outa09ol-DFC_rbr_outA09OL.st ---- *)
(* --- Interface --- *)
{attribute 'external_name' := 'cmp_rts_DFC_rbr_outA09OL'}
TYPE DFC_rbr_outA09OL :
STRUCT
	DTC: UDINT := 16#142B00;
	DFCid: UINT := 303;
	debounceMethod: USINT := TIME_UP_DOWN;
END_STRUCT
END_TYPE

(* ---- dfc_rbr_outa09or-DFC_rbr_outA09OR.st ---- *)
(* --- Interface --- *)
{attribute 'external_name' := 'cmp_rts_DFC_rbr_outA09OR'}
TYPE DFC_rbr_outA09OR :
STRUCT
	DTC: UDINT := 16#142C00;
	DFCid: UINT := 304;
	debounceMethod: USINT := TIME_UP_DOWN;
END_STRUCT
END_TYPE
